Yaskawa INFORM job: 4043MM.JBI

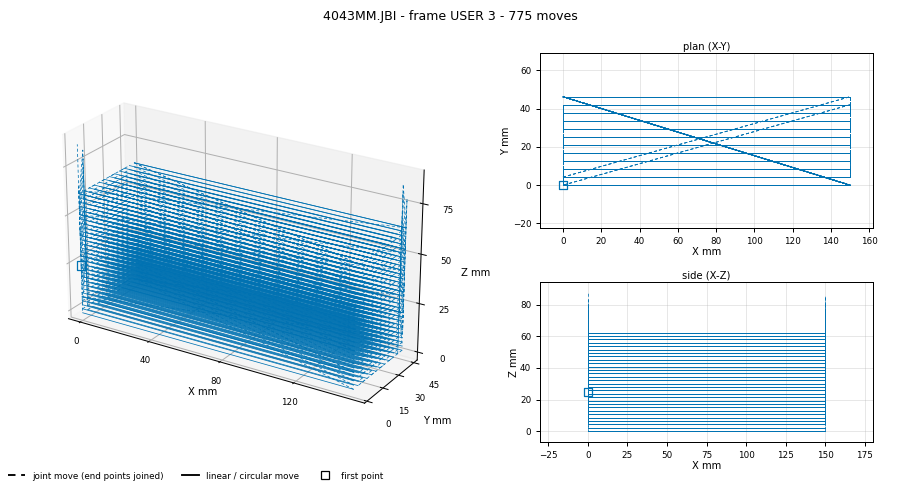
[picture p0: tool path of 4043MM.JBI in frame USER 3, 775 of 775 moves have a stored position in this frame; points joined in program order, loops and branches not executed]
/JOB
//NAME 4043MM
//POS
///NPOS 775,0,0,0,0,0
///USER 3
///TOOL 1
///POSTYPE USER
///RECTAN
///RCONF 1,0,0,0,0,0,0,0,0,0,0,0,0,0,0,0,0,0,0,0,0,0,0,0
C00000=0.000,0.000,25.000,0.0000,0.0000,-110.0000
C00001=0.000,0.000,0.000,0.0000,0.0000,-110.0000
C00002=150.000,0.000,0.000,0.0000,0.0000,-110.0000
C00003=0.000,46.200,0.000,0.0000,0.0000,-110.0000
C00004=150.000,46.200,0.000,0.0000,0.0000,-110.0000
C00005=150.000,4.200,0.000,0.0000,0.0000,-110.0000
C00006=0.000,4.200,0.000,0.0000,0.0000,-110.0000
C00007=0.000,8.400,0.000,0.0000,0.0000,-110.0000
C00008=150.000,8.400,0.000,0.0000,0.0000,-110.0000
C00009=150.000,12.600,0.000,0.0000,0.0000,-110.0000
C00010=0.000,12.600,0.000,0.0000,0.0000,-110.0000
C00011=0.000,16.800,0.000,0.0000,0.0000,-110.0000
C00012=150.000,16.800,0.000,0.0000,0.0000,-110.0000
C00013=150.000,21.000,0.000,0.0000,0.0000,-110.0000
C00014=0.000,21.000,0.000,0.0000,0.0000,-110.0000
C00015=0.000,25.200,0.000,0.0000,0.0000,-110.0000
C00016=150.000,25.200,0.000,0.0000,0.0000,-110.0000
C00017=150.000,29.400,0.000,0.0000,0.0000,-110.0000
C00018=0.000,29.400,0.000,0.0000,0.0000,-110.0000
C00019=0.000,33.600,0.000,0.0000,0.0000,-110.0000
C00020=150.000,33.600,0.000,0.0000,0.0000,-110.0000
C00021=150.000,37.800,0.000,0.0000,0.0000,-110.0000
C00022=0.000,37.800,0.000,0.0000,0.0000,-110.0000
C00023=0.000,42.000,0.000,0.0000,0.0000,-110.0000
C00024=150.000,42.000,0.000,0.0000,0.0000,-110.0000
C00025=150.000,42.000,25.000,0.0000,0.0000,-110.0000
C00026=150.000,46.200,2.150,0.0000,0.0000,-110.0000
C00027=0.000,46.200,2.150,0.0000,0.0000,-110.0000
C00028=150.000,0.000,2.150,0.0000,0.0000,-110.0000
C00029=0.000,0.000,2.150,0.0000,0.0000,-110.0000
C00030=0.000,42.000,2.150,0.0000,0.0000,-110.0000
C00031=150.000,42.000,2.150,0.0000,0.0000,-110.0000
C00032=150.000,37.800,2.150,0.0000,0.0000,-110.0000
C00033=0.000,37.800,2.150,0.0000,0.0000,-110.0000
C00034=0.000,33.600,2.150,0.0000,0.0000,-110.0000
C00035=150.000,33.600,2.150,0.0000,0.0000,-110.0000
C00036=150.000,29.400,2.150,0.0000,0.0000,-110.0000
C00037=0.000,29.400,2.150,0.0000,0.0000,-110.0000
C00038=0.000,25.200,2.150,0.0000,0.0000,-110.0000
C00039=150.000,25.200,2.150,0.0000,0.0000,-110.0000
C00040=150.000,21.000,2.150,0.0000,0.0000,-110.0000
C00041=0.000,21.000,2.150,0.0000,0.0000,-110.0000
C00042=0.000,16.800,2.150,0.0000,0.0000,-110.0000
C00043=150.000,16.800,2.150,0.0000,0.0000,-110.0000
C00044=150.000,12.600,2.150,0.0000,0.0000,-110.0000
C00045=0.000,12.600,2.150,0.0000,0.0000,-110.0000
C00046=0.000,8.400,2.150,0.0000,0.0000,-110.0000
C00047=150.000,8.400,2.150,0.0000,0.0000,-110.0000
C00048=150.000,4.200,2.150,0.0000,0.0000,-110.0000
C00049=0.000,4.200,2.150,0.0000,0.0000,-110.0000
C00050=0.000,4.200,27.150,0.0000,0.0000,-110.0000
C00051=0.000,0.000,4.300,0.0000,0.0000,-110.0000
C00052=150.000,0.000,4.300,0.0000,0.0000,-110.0000
C00053=0.000,46.200,4.300,0.0000,0.0000,-110.0000
C00054=150.000,46.200,4.300,0.0000,0.0000,-110.0000
C00055=150.000,4.200,4.300,0.0000,0.0000,-110.0000
C00056=0.000,4.200,4.300,0.0000,0.0000,-110.0000
C00057=0.000,8.400,4.300,0.0000,0.0000,-110.0000
C00058=150.000,8.400,4.300,0.0000,0.0000,-110.0000
C00059=150.000,12.600,4.300,0.0000,0.0000,-110.0000
C00060=0.000,12.600,4.300,0.0000,0.0000,-110.0000
C00061=0.000,16.800,4.300,0.0000,0.0000,-110.0000
C00062=150.000,16.800,4.300,0.0000,0.0000,-110.0000
C00063=150.000,21.000,4.300,0.0000,0.0000,-110.0000
C00064=0.000,21.000,4.300,0.0000,0.0000,-110.0000
C00065=0.000,25.200,4.300,0.0000,0.0000,-110.0000
C00066=150.000,25.200,4.300,0.0000,0.0000,-110.0000
C00067=150.000,29.400,4.300,0.0000,0.0000,-110.0000
C00068=0.000,29.400,4.300,0.0000,0.0000,-110.0000
C00069=0.000,33.600,4.300,0.0000,0.0000,-110.0000
C00070=150.000,33.600,4.300,0.0000,0.0000,-110.0000
C00071=150.000,37.800,4.300,0.0000,0.0000,-110.0000
C00072=0.000,37.800,4.300,0.0000,0.0000,-110.0000
C00073=0.000,42.000,4.300,0.0000,0.0000,-110.0000
C00074=150.000,42.000,4.300,0.0000,0.0000,-110.0000
C00075=150.000,42.000,29.300,0.0000,0.0000,-110.0000
C00076=150.000,46.200,6.450,0.0000,0.0000,-110.0000
C00077=0.000,46.200,6.450,0.0000,0.0000,-110.0000
C00078=150.000,0.000,6.450,0.0000,0.0000,-110.0000
C00079=0.000,0.000,6.450,0.0000,0.0000,-110.0000
C00080=0.000,42.000,6.450,0.0000,0.0000,-110.0000
C00081=150.000,42.000,6.450,0.0000,0.0000,-110.0000
C00082=150.000,37.800,6.450,0.0000,0.0000,-110.0000
C00083=0.000,37.800,6.450,0.0000,0.0000,-110.0000
C00084=0.000,33.600,6.450,0.0000,0.0000,-110.0000
C00085=150.000,33.600,6.450,0.0000,0.0000,-110.0000
C00086=150.000,29.400,6.450,0.0000,0.0000,-110.0000
C00087=0.000,29.400,6.450,0.0000,0.0000,-110.0000
C00088=0.000,25.200,6.450,0.0000,0.0000,-110.0000
C00089=150.000,25.200,6.450,0.0000,0.0000,-110.0000
C00090=150.000,21.000,6.450,0.0000,0.0000,-110.0000
C00091=0.000,21.000,6.450,0.0000,0.0000,-110.0000
C00092=0.000,16.800,6.450,0.0000,0.0000,-110.0000
C00093=150.000,16.800,6.450,0.0000,0.0000,-110.0000
C00094=150.000,12.600,6.450,0.0000,0.0000,-110.0000
C00095=0.000,12.600,6.450,0.0000,0.0000,-110.0000
C00096=0.000,8.400,6.450,0.0000,0.0000,-110.0000
C00097=150.000,8.400,6.450,0.0000,0.0000,-110.0000
C00098=150.000,4.200,6.450,0.0000,0.0000,-110.0000
C00099=0.000,4.200,6.450,0.0000,0.0000,-110.0000
C00100=0.000,4.200,31.450,0.0000,0.0000,-110.0000
C00101=0.000,0.000,8.600,0.0000,0.0000,-110.0000
C00102=150.000,0.000,8.600,0.0000,0.0000,-110.0000
C00103=0.000,46.200,8.600,0.0000,0.0000,-110.0000
C00104=150.000,46.200,8.600,0.0000,0.0000,-110.0000
C00105=150.000,4.200,8.600,0.0000,0.0000,-110.0000
C00106=0.000,4.200,8.600,0.0000,0.0000,-110.0000
C00107=0.000,8.400,8.600,0.0000,0.0000,-110.0000
C00108=150.000,8.400,8.600,0.0000,0.0000,-110.0000
C00109=150.000,12.600,8.600,0.0000,0.0000,-110.0000
C00110=0.000,12.600,8.600,0.0000,0.0000,-110.0000
C00111=0.000,16.800,8.600,0.0000,0.0000,-110.0000
C00112=150.000,16.800,8.600,0.0000,0.0000,-110.0000
C00113=150.000,21.000,8.600,0.0000,0.0000,-110.0000
C00114=0.000,21.000,8.600,0.0000,0.0000,-110.0000
C00115=0.000,25.200,8.600,0.0000,0.0000,-110.0000
C00116=150.000,25.200,8.600,0.0000,0.0000,-110.0000
C00117=150.000,29.400,8.600,0.0000,0.0000,-110.0000
C00118=0.000,29.400,8.600,0.0000,0.0000,-110.0000
C00119=0.000,33.600,8.600,0.0000,0.0000,-110.0000
C00120=150.000,33.600,8.600,0.0000,0.0000,-110.0000
C00121=150.000,37.800,8.600,0.0000,0.0000,-110.0000
C00122=0.000,37.800,8.600,0.0000,0.0000,-110.0000
C00123=0.000,42.000,8.600,0.0000,0.0000,-110.0000
C00124=150.000,42.000,8.600,0.0000,0.0000,-110.0000
C00125=0.000,0.000,8.600,0.0000,0.0000,-110.0000
C00126=150.000,0.000,8.600,0.0000,0.0000,-110.0000
C00127=0.000,46.200,8.600,0.0000,0.0000,-110.0000
C00128=150.000,46.200,8.600,0.0000,0.0000,-110.0000
C00129=150.000,46.200,33.600,0.0000,0.0000,-110.0000
C00130=150.000,46.200,10.750,0.0000,0.0000,-110.0000
C00131=0.000,46.200,10.750,0.0000,0.0000,-110.0000
C00132=150.000,0.000,10.750,0.0000,0.0000,-110.0000
C00133=0.000,0.000,10.750,0.0000,0.0000,-110.0000
C00134=0.000,42.000,10.750,0.0000,0.0000,-110.0000
C00135=150.000,42.000,10.750,0.0000,0.0000,-110.0000
C00136=150.000,37.800,10.750,0.0000,0.0000,-110.0000
C00137=0.000,37.800,10.750,0.0000,0.0000,-110.0000
C00138=0.000,33.600,10.750,0.0000,0.0000,-110.0000
C00139=150.000,33.600,10.750,0.0000,0.0000,-110.0000
C00140=150.000,29.400,10.750,0.0000,0.0000,-110.0000
C00141=0.000,29.400,10.750,0.0000,0.0000,-110.0000
C00142=0.000,25.200,10.750,0.0000,0.0000,-110.0000
C00143=150.000,25.200,10.750,0.0000,0.0000,-110.0000
C00144=150.000,21.000,10.750,0.0000,0.0000,-110.0000
C00145=0.000,21.000,10.750,0.0000,0.0000,-110.0000
C00146=0.000,16.800,10.750,0.0000,0.0000,-110.0000
C00147=150.000,16.800,10.750,0.0000,0.0000,-110.0000
C00148=150.000,12.600,10.750,0.0000,0.0000,-110.0000
C00149=0.000,12.600,10.750,0.0000,0.0000,-110.0000
C00150=0.000,8.400,10.750,0.0000,0.0000,-110.0000
C00151=150.000,8.400,10.750,0.0000,0.0000,-110.0000
C00152=150.000,4.200,10.750,0.0000,0.0000,-110.0000
C00153=0.000,4.200,10.750,0.0000,0.0000,-110.0000
C00154=0.000,4.200,35.750,0.0000,0.0000,-110.0000
C00155=0.000,0.000,12.900,0.0000,0.0000,-110.0000
C00156=150.000,0.000,12.900,0.0000,0.0000,-110.0000
C00157=0.000,46.200,12.900,0.0000,0.0000,-110.0000
C00158=150.000,46.200,12.900,0.0000,0.0000,-110.0000
C00159=150.000,4.200,12.900,0.0000,0.0000,-110.0000
C00160=0.000,4.200,12.900,0.0000,0.0000,-110.0000
C00161=0.000,8.400,12.900,0.0000,0.0000,-110.0000
C00162=150.000,8.400,12.900,0.0000,0.0000,-110.0000
C00163=150.000,12.600,12.900,0.0000,0.0000,-110.0000
C00164=0.000,12.600,12.900,0.0000,0.0000,-110.0000
C00165=0.000,16.800,12.900,0.0000,0.0000,-110.0000
C00166=150.000,16.800,12.900,0.0000,0.0000,-110.0000
C00167=150.000,21.000,12.900,0.0000,0.0000,-110.0000
C00168=0.000,21.000,12.900,0.0000,0.0000,-110.0000
C00169=0.000,25.200,12.900,0.0000,0.0000,-110.0000
C00170=150.000,25.200,12.900,0.0000,0.0000,-110.0000
C00171=150.000,29.400,12.900,0.0000,0.0000,-110.0000
C00172=0.000,29.400,12.900,0.0000,0.0000,-110.0000
C00173=0.000,33.600,12.900,0.0000,0.0000,-110.0000
C00174=150.000,33.600,12.900,0.0000,0.0000,-110.0000
C00175=150.000,37.800,12.900,0.0000,0.0000,-110.0000
C00176=0.000,37.800,12.900,0.0000,0.0000,-110.0000
C00177=0.000,42.000,12.900,0.0000,0.0000,-110.0000
C00178=150.000,42.000,12.900,0.0000,0.0000,-110.0000
C00179=150.000,42.000,37.900,0.0000,0.0000,-110.0000
C00180=150.000,46.200,15.050,0.0000,0.0000,-110.0000
C00181=0.000,46.200,15.050,0.0000,0.0000,-110.0000
C00182=150.000,0.000,15.050,0.0000,0.0000,-110.0000
C00183=0.000,0.000,15.050,0.0000,0.0000,-110.0000
C00184=0.000,42.000,15.050,0.0000,0.0000,-110.0000
C00185=150.000,42.000,15.050,0.0000,0.0000,-110.0000
C00186=150.000,37.800,15.050,0.0000,0.0000,-110.0000
C00187=0.000,37.800,15.050,0.0000,0.0000,-110.0000
C00188=0.000,33.600,15.050,0.0000,0.0000,-110.0000
C00189=150.000,33.600,15.050,0.0000,0.0000,-110.0000
C00190=150.000,29.400,15.050,0.0000,0.0000,-110.0000
C00191=0.000,29.400,15.050,0.0000,0.0000,-110.0000
C00192=0.000,25.200,15.050,0.0000,0.0000,-110.0000
C00193=150.000,25.200,15.050,0.0000,0.0000,-110.0000
C00194=150.000,21.000,15.050,0.0000,0.0000,-110.0000
C00195=0.000,21.000,15.050,0.0000,0.0000,-110.0000
C00196=0.000,16.800,15.050,0.0000,0.0000,-110.0000
C00197=150.000,16.800,15.050,0.0000,0.0000,-110.0000
C00198=150.000,12.600,15.050,0.0000,0.0000,-110.0000
C00199=0.000,12.600,15.050,0.0000,0.0000,-110.0000
C00200=0.000,8.400,15.050,0.0000,0.0000,-110.0000
C00201=150.000,8.400,15.050,0.0000,0.0000,-110.0000
C00202=150.000,4.200,15.050,0.0000,0.0000,-110.0000
C00203=0.000,4.200,15.050,0.0000,0.0000,-110.0000
C00204=0.000,4.200,40.050,0.0000,0.0000,-110.0000
C00205=0.000,0.000,17.200,0.0000,0.0000,-110.0000
C00206=150.000,0.000,17.200,0.0000,0.0000,-110.0000
C00207=0.000,46.200,17.200,0.0000,0.0000,-110.0000
C00208=150.000,46.200,17.200,0.0000,0.0000,-110.0000
C00209=150.000,4.200,17.200,0.0000,0.0000,-110.0000
C00210=0.000,4.200,17.200,0.0000,0.0000,-110.0000
C00211=0.000,8.400,17.200,0.0000,0.0000,-110.0000
C00212=150.000,8.400,17.200,0.0000,0.0000,-110.0000
C00213=150.000,12.600,17.200,0.0000,0.0000,-110.0000
C00214=0.000,12.600,17.200,0.0000,0.0000,-110.0000
C00215=0.000,16.800,17.200,0.0000,0.0000,-110.0000
C00216=150.000,16.800,17.200,0.0000,0.0000,-110.0000
C00217=150.000,21.000,17.200,0.0000,0.0000,-110.0000
C00218=0.000,21.000,17.200,0.0000,0.0000,-110.0000
C00219=0.000,25.200,17.200,0.0000,0.0000,-110.0000
C00220=150.000,25.200,17.200,0.0000,0.0000,-110.0000
C00221=150.000,29.400,17.200,0.0000,0.0000,-110.0000
C00222=0.000,29.400,17.200,0.0000,0.0000,-110.0000
C00223=0.000,33.600,17.200,0.0000,0.0000,-110.0000
C00224=150.000,33.600,17.200,0.0000,0.0000,-110.0000
C00225=150.000,37.800,17.200,0.0000,0.0000,-110.0000
C00226=0.000,37.800,17.200,0.0000,0.0000,-110.0000
C00227=0.000,42.000,17.200,0.0000,0.0000,-110.0000
C00228=150.000,42.000,17.200,0.0000,0.0000,-110.0000
C00229=150.000,42.000,42.200,0.0000,0.0000,-110.0000
C00230=150.000,46.200,19.350,0.0000,0.0000,-110.0000
C00231=0.000,46.200,19.350,0.0000,0.0000,-110.0000
C00232=150.000,0.000,19.350,0.0000,0.0000,-110.0000
C00233=0.000,0.000,19.350,0.0000,0.0000,-110.0000
C00234=0.000,42.000,19.350,0.0000,0.0000,-110.0000
C00235=150.000,42.000,19.350,0.0000,0.0000,-110.0000
C00236=150.000,37.800,19.350,0.0000,0.0000,-110.0000
C00237=0.000,37.800,19.350,0.0000,0.0000,-110.0000
C00238=0.000,33.600,19.350,0.0000,0.0000,-110.0000
C00239=150.000,33.600,19.350,0.0000,0.0000,-110.0000
C00240=150.000,29.400,19.350,0.0000,0.0000,-110.0000
C00241=0.000,29.400,19.350,0.0000,0.0000,-110.0000
C00242=0.000,25.200,19.350,0.0000,0.0000,-110.0000
C00243=150.000,25.200,19.350,0.0000,0.0000,-110.0000
C00244=150.000,21.000,19.350,0.0000,0.0000,-110.0000
C00245=0.000,21.000,19.350,0.0000,0.0000,-110.0000
C00246=0.000,16.800,19.350,0.0000,0.0000,-110.0000
C00247=150.000,16.800,19.350,0.0000,0.0000,-110.0000
C00248=150.000,12.600,19.350,0.0000,0.0000,-110.0000
C00249=0.000,12.600,19.350,0.0000,0.0000,-110.0000
C00250=0.000,8.400,19.350,0.0000,0.0000,-110.0000
C00251=150.000,8.400,19.350,0.0000,0.0000,-110.0000
C00252=150.000,4.200,19.350,0.0000,0.0000,-110.0000
C00253=0.000,4.200,19.350,0.0000,0.0000,-110.0000
C00254=150.000,46.200,19.350,0.0000,0.0000,-110.0000
C00255=0.000,46.200,19.350,0.0000,0.0000,-110.0000
C00256=150.000,0.000,19.350,0.0000,0.0000,-110.0000
C00257=0.000,0.000,19.350,0.0000,0.0000,-110.0000
C00258=0.000,0.000,44.350,0.0000,0.0000,-110.0000
C00259=0.000,0.000,21.500,0.0000,0.0000,-110.0000
C00260=150.000,0.000,21.500,0.0000,0.0000,-110.0000
C00261=0.000,46.200,21.500,0.0000,0.0000,-110.0000
C00262=150.000,46.200,21.500,0.0000,0.0000,-110.0000
C00263=150.000,4.200,21.500,0.0000,0.0000,-110.0000
C00264=0.000,4.200,21.500,0.0000,0.0000,-110.0000
C00265=0.000,8.400,21.500,0.0000,0.0000,-110.0000
C00266=150.000,8.400,21.500,0.0000,0.0000,-110.0000
C00267=150.000,12.600,21.500,0.0000,0.0000,-110.0000
C00268=0.000,12.600,21.500,0.0000,0.0000,-110.0000
C00269=0.000,16.800,21.500,0.0000,0.0000,-110.0000
C00270=150.000,16.800,21.500,0.0000,0.0000,-110.0000
C00271=150.000,21.000,21.500,0.0000,0.0000,-110.0000
C00272=0.000,21.000,21.500,0.0000,0.0000,-110.0000
C00273=0.000,25.200,21.500,0.0000,0.0000,-110.0000
C00274=150.000,25.200,21.500,0.0000,0.0000,-110.0000
C00275=150.000,29.400,21.500,0.0000,0.0000,-110.0000
C00276=0.000,29.400,21.500,0.0000,0.0000,-110.0000
C00277=0.000,33.600,21.500,0.0000,0.0000,-110.0000
C00278=150.000,33.600,21.500,0.0000,0.0000,-110.0000
C00279=150.000,37.800,21.500,0.0000,0.0000,-110.0000
C00280=0.000,37.800,21.500,0.0000,0.0000,-110.0000
C00281=0.000,42.000,21.500,0.0000,0.0000,-110.0000
C00282=150.000,42.000,21.500,0.0000,0.0000,-110.0000
C00283=150.000,42.000,46.500,0.0000,0.0000,-110.0000
C00284=150.000,46.200,23.650,0.0000,0.0000,-110.0000
C00285=0.000,46.200,23.650,0.0000,0.0000,-110.0000
C00286=150.000,0.000,23.650,0.0000,0.0000,-110.0000
C00287=0.000,0.000,23.650,0.0000,0.0000,-110.0000
C00288=0.000,42.000,23.650,0.0000,0.0000,-110.0000
C00289=150.000,42.000,23.650,0.0000,0.0000,-110.0000
C00290=150.000,37.800,23.650,0.0000,0.0000,-110.0000
C00291=0.000,37.800,23.650,0.0000,0.0000,-110.0000
C00292=0.000,33.600,23.650,0.0000,0.0000,-110.0000
C00293=150.000,33.600,23.650,0.0000,0.0000,-110.0000
C00294=150.000,29.400,23.650,0.0000,0.0000,-110.0000
C00295=0.000,29.400,23.650,0.0000,0.0000,-110.0000
C00296=0.000,25.200,23.650,0.0000,0.0000,-110.0000
C00297=150.000,25.200,23.650,0.0000,0.0000,-110.0000
C00298=150.000,21.000,23.650,0.0000,0.0000,-110.0000
C00299=0.000,21.000,23.650,0.0000,0.0000,-110.0000
C00300=0.000,16.800,23.650,0.0000,0.0000,-110.0000
C00301=150.000,16.800,23.650,0.0000,0.0000,-110.0000
C00302=150.000,12.600,23.650,0.0000,0.0000,-110.0000
C00303=0.000,12.600,23.650,0.0000,0.0000,-110.0000
C00304=0.000,8.400,23.650,0.0000,0.0000,-110.0000
C00305=150.000,8.400,23.650,0.0000,0.0000,-110.0000
C00306=150.000,4.200,23.650,0.0000,0.0000,-110.0000
C00307=0.000,4.200,23.650,0.0000,0.0000,-110.0000
C00308=0.000,4.200,48.650,0.0000,0.0000,-110.0000
C00309=0.000,0.000,25.800,0.0000,0.0000,-110.0000
C00310=150.000,0.000,25.800,0.0000,0.0000,-110.0000
C00311=0.000,46.200,25.800,0.0000,0.0000,-110.0000
C00312=150.000,46.200,25.800,0.0000,0.0000,-110.0000
C00313=150.000,4.200,25.800,0.0000,0.0000,-110.0000
C00314=0.000,4.200,25.800,0.0000,0.0000,-110.0000
C00315=0.000,8.400,25.800,0.0000,0.0000,-110.0000
C00316=150.000,8.400,25.800,0.0000,0.0000,-110.0000
C00317=150.000,12.600,25.800,0.0000,0.0000,-110.0000
C00318=0.000,12.600,25.800,0.0000,0.0000,-110.0000
C00319=0.000,16.800,25.800,0.0000,0.0000,-110.0000
C00320=150.000,16.800,25.800,0.0000,0.0000,-110.0000
C00321=150.000,21.000,25.800,0.0000,0.0000,-110.0000
C00322=0.000,21.000,25.800,0.0000,0.0000,-110.0000
C00323=0.000,25.200,25.800,0.0000,0.0000,-110.0000
C00324=150.000,25.200,25.800,0.0000,0.0000,-110.0000
C00325=150.000,29.400,25.800,0.0000,0.0000,-110.0000
C00326=0.000,29.400,25.800,0.0000,0.0000,-110.0000
C00327=0.000,33.600,25.800,0.0000,0.0000,-110.0000
C00328=150.000,33.600,25.800,0.0000,0.0000,-110.0000
C00329=150.000,37.800,25.800,0.0000,0.0000,-110.0000
C00330=0.000,37.800,25.800,0.0000,0.0000,-110.0000
C00331=0.000,42.000,25.800,0.0000,0.0000,-110.0000
C00332=150.000,42.000,25.800,0.0000,0.0000,-110.0000
C00333=150.000,42.000,50.800,0.0000,0.0000,-110.0000
C00334=150.000,46.200,27.950,0.0000,0.0000,-110.0000
C00335=0.000,46.200,27.950,0.0000,0.0000,-110.0000
C00336=150.000,0.000,27.950,0.0000,0.0000,-110.0000
C00337=0.000,0.000,27.950,0.0000,0.0000,-110.0000
C00338=0.000,42.000,27.950,0.0000,0.0000,-110.0000
C00339=150.000,42.000,27.950,0.0000,0.0000,-110.0000
C00340=150.000,37.800,27.950,0.0000,0.0000,-110.0000
C00341=0.000,37.800,27.950,0.0000,0.0000,-110.0000
C00342=0.000,33.600,27.950,0.0000,0.0000,-110.0000
C00343=150.000,33.600,27.950,0.0000,0.0000,-110.0000
C00344=150.000,29.400,27.950,0.0000,0.0000,-110.0000
C00345=0.000,29.400,27.950,0.0000,0.0000,-110.0000
C00346=0.000,25.200,27.950,0.0000,0.0000,-110.0000
C00347=150.000,25.200,27.950,0.0000,0.0000,-110.0000
C00348=150.000,21.000,27.950,0.0000,0.0000,-110.0000
C00349=0.000,21.000,27.950,0.0000,0.0000,-110.0000
C00350=0.000,16.800,27.950,0.0000,0.0000,-110.0000
C00351=150.000,16.800,27.950,0.0000,0.0000,-110.0000
C00352=150.000,12.600,27.950,0.0000,0.0000,-110.0000
C00353=0.000,12.600,27.950,0.0000,0.0000,-110.0000
C00354=0.000,8.400,27.950,0.0000,0.0000,-110.0000
C00355=150.000,8.400,27.950,0.0000,0.0000,-110.0000
C00356=150.000,4.200,27.950,0.0000,0.0000,-110.0000
C00357=0.000,4.200,27.950,0.0000,0.0000,-110.0000
C00358=0.000,4.200,52.950,0.0000,0.0000,-110.0000
C00359=0.000,0.000,30.100,0.0000,0.0000,-110.0000
C00360=150.000,0.000,30.100,0.0000,0.0000,-110.0000
C00361=0.000,46.200,30.100,0.0000,0.0000,-110.0000
C00362=150.000,46.200,30.100,0.0000,0.0000,-110.0000
C00363=150.000,4.200,30.100,0.0000,0.0000,-110.0000
C00364=0.000,4.200,30.100,0.0000,0.0000,-110.0000
C00365=0.000,8.400,30.100,0.0000,0.0000,-110.0000
C00366=150.000,8.400,30.100,0.0000,0.0000,-110.0000
C00367=150.000,12.600,30.100,0.0000,0.0000,-110.0000
C00368=0.000,12.600,30.100,0.0000,0.0000,-110.0000
C00369=0.000,16.800,30.100,0.0000,0.0000,-110.0000
C00370=150.000,16.800,30.100,0.0000,0.0000,-110.0000
C00371=150.000,21.000,30.100,0.0000,0.0000,-110.0000
C00372=0.000,21.000,30.100,0.0000,0.0000,-110.0000
C00373=0.000,25.200,30.100,0.0000,0.0000,-110.0000
C00374=150.000,25.200,30.100,0.0000,0.0000,-110.0000
C00375=150.000,29.400,30.100,0.0000,0.0000,-110.0000
C00376=0.000,29.400,30.100,0.0000,0.0000,-110.0000
C00377=0.000,33.600,30.100,0.0000,0.0000,-110.0000
C00378=150.000,33.600,30.100,0.0000,0.0000,-110.0000
C00379=150.000,37.800,30.100,0.0000,0.0000,-110.0000
C00380=0.000,37.800,30.100,0.0000,0.0000,-110.0000
C00381=0.000,42.000,30.100,0.0000,0.0000,-110.0000
C00382=150.000,42.000,30.100,0.0000,0.0000,-110.0000
C00383=0.000,0.000,30.100,0.0000,0.0000,-110.0000
C00384=150.000,0.000,30.100,0.0000,0.0000,-110.0000
C00385=0.000,46.200,30.100,0.0000,0.0000,-110.0000
C00386=150.000,46.200,30.100,0.0000,0.0000,-110.0000
C00387=150.000,46.200,55.100,0.0000,0.0000,-110.0000
C00388=150.000,46.200,32.250,0.0000,0.0000,-110.0000
C00389=0.000,46.200,32.250,0.0000,0.0000,-110.0000
C00390=150.000,0.000,32.250,0.0000,0.0000,-110.0000
C00391=0.000,0.000,32.250,0.0000,0.0000,-110.0000
C00392=0.000,42.000,32.250,0.0000,0.0000,-110.0000
C00393=150.000,42.000,32.250,0.0000,0.0000,-110.0000
C00394=150.000,37.800,32.250,0.0000,0.0000,-110.0000
C00395=0.000,37.800,32.250,0.0000,0.0000,-110.0000
C00396=0.000,33.600,32.250,0.0000,0.0000,-110.0000
C00397=150.000,33.600,32.250,0.0000,0.0000,-110.0000
C00398=150.000,29.400,32.250,0.0000,0.0000,-110.0000
C00399=0.000,29.400,32.250,0.0000,0.0000,-110.0000
C00400=0.000,25.200,32.250,0.0000,0.0000,-110.0000
C00401=150.000,25.200,32.250,0.0000,0.0000,-110.0000
C00402=150.000,21.000,32.250,0.0000,0.0000,-110.0000
C00403=0.000,21.000,32.250,0.0000,0.0000,-110.0000
C00404=0.000,16.800,32.250,0.0000,0.0000,-110.0000
C00405=150.000,16.800,32.250,0.0000,0.0000,-110.0000
C00406=150.000,12.600,32.250,0.0000,0.0000,-110.0000
C00407=0.000,12.600,32.250,0.0000,0.0000,-110.0000
C00408=0.000,8.400,32.250,0.0000,0.0000,-110.0000
C00409=150.000,8.400,32.250,0.0000,0.0000,-110.0000
C00410=150.000,4.200,32.250,0.0000,0.0000,-110.0000
C00411=0.000,4.200,32.250,0.0000,0.0000,-110.0000
C00412=0.000,4.200,57.250,0.0000,0.0000,-110.0000
C00413=0.000,0.000,34.400,0.0000,0.0000,-110.0000
C00414=150.000,0.000,34.400,0.0000,0.0000,-110.0000
C00415=0.000,46.200,34.400,0.0000,0.0000,-110.0000
C00416=150.000,46.200,34.400,0.0000,0.0000,-110.0000
C00417=150.000,4.200,34.400,0.0000,0.0000,-110.0000
C00418=0.000,4.200,34.400,0.0000,0.0000,-110.0000
C00419=0.000,8.400,34.400,0.0000,0.0000,-110.0000
C00420=150.000,8.400,34.400,0.0000,0.0000,-110.0000
C00421=150.000,12.600,34.400,0.0000,0.0000,-110.0000
C00422=0.000,12.600,34.400,0.0000,0.0000,-110.0000
C00423=0.000,16.800,34.400,0.0000,0.0000,-110.0000
C00424=150.000,16.800,34.400,0.0000,0.0000,-110.0000
C00425=150.000,21.000,34.400,0.0000,0.0000,-110.0000
C00426=0.000,21.000,34.400,0.0000,0.0000,-110.0000
C00427=0.000,25.200,34.400,0.0000,0.0000,-110.0000
C00428=150.000,25.200,34.400,0.0000,0.0000,-110.0000
C00429=150.000,29.400,34.400,0.0000,0.0000,-110.0000
C00430=0.000,29.400,34.400,0.0000,0.0000,-110.0000
C00431=0.000,33.600,34.400,0.0000,0.0000,-110.0000
C00432=150.000,33.600,34.400,0.0000,0.0000,-110.0000
C00433=150.000,37.800,34.400,0.0000,0.0000,-110.0000
C00434=0.000,37.800,34.400,0.0000,0.0000,-110.0000
C00435=0.000,42.000,34.400,0.0000,0.0000,-110.0000
C00436=150.000,42.000,34.400,0.0000,0.0000,-110.0000
C00437=150.000,42.000,59.400,0.0000,0.0000,-110.0000
C00438=150.000,46.200,36.550,0.0000,0.0000,-110.0000
C00439=0.000,46.200,36.550,0.0000,0.0000,-110.0000
C00440=150.000,0.000,36.550,0.0000,0.0000,-110.0000
C00441=0.000,0.000,36.550,0.0000,0.0000,-110.0000
C00442=0.000,42.000,36.550,0.0000,0.0000,-110.0000
C00443=150.000,42.000,36.550,0.0000,0.0000,-110.0000
C00444=150.000,37.800,36.550,0.0000,0.0000,-110.0000
C00445=0.000,37.800,36.550,0.0000,0.0000,-110.0000
C00446=0.000,33.600,36.550,0.0000,0.0000,-110.0000
C00447=150.000,33.600,36.550,0.0000,0.0000,-110.0000
C00448=150.000,29.400,36.550,0.0000,0.0000,-110.0000
C00449=0.000,29.400,36.550,0.0000,0.0000,-110.0000
C00450=0.000,25.200,36.550,0.0000,0.0000,-110.0000
C00451=150.000,25.200,36.550,0.0000,0.0000,-110.0000
C00452=150.000,21.000,36.550,0.0000,0.0000,-110.0000
C00453=0.000,21.000,36.550,0.0000,0.0000,-110.0000
C00454=0.000,16.800,36.550,0.0000,0.0000,-110.0000
C00455=150.000,16.800,36.550,0.0000,0.0000,-110.0000
C00456=150.000,12.600,36.550,0.0000,0.0000,-110.0000
C00457=0.000,12.600,36.550,0.0000,0.0000,-110.0000
C00458=0.000,8.400,36.550,0.0000,0.0000,-110.0000
C00459=150.000,8.400,36.550,0.0000,0.0000,-110.0000
C00460=150.000,4.200,36.550,0.0000,0.0000,-110.0000
C00461=0.000,4.200,36.550,0.0000,0.0000,-110.0000
C00462=0.000,4.200,61.550,0.0000,0.0000,-110.0000
C00463=0.000,0.000,38.700,0.0000,0.0000,-110.0000
C00464=150.000,0.000,38.700,0.0000,0.0000,-110.0000
C00465=0.000,46.200,38.700,0.0000,0.0000,-110.0000
C00466=150.000,46.200,38.700,0.0000,0.0000,-110.0000
C00467=150.000,4.200,38.700,0.0000,0.0000,-110.0000
C00468=0.000,4.200,38.700,0.0000,0.0000,-110.0000
C00469=0.000,8.400,38.700,0.0000,0.0000,-110.0000
C00470=150.000,8.400,38.700,0.0000,0.0000,-110.0000
C00471=150.000,12.600,38.700,0.0000,0.0000,-110.0000
C00472=0.000,12.600,38.700,0.0000,0.0000,-110.0000
C00473=0.000,16.800,38.700,0.0000,0.0000,-110.0000
C00474=150.000,16.800,38.700,0.0000,0.0000,-110.0000
C00475=150.000,21.000,38.700,0.0000,0.0000,-110.0000
C00476=0.000,21.000,38.700,0.0000,0.0000,-110.0000
C00477=0.000,25.200,38.700,0.0000,0.0000,-110.0000
C00478=150.000,25.200,38.700,0.0000,0.0000,-110.0000
C00479=150.000,29.400,38.700,0.0000,0.0000,-110.0000
C00480=0.000,29.400,38.700,0.0000,0.0000,-110.0000
C00481=0.000,33.600,38.700,0.0000,0.0000,-110.0000
C00482=150.000,33.600,38.700,0.0000,0.0000,-110.0000
C00483=150.000,37.800,38.700,0.0000,0.0000,-110.0000
C00484=0.000,37.800,38.700,0.0000,0.0000,-110.0000
C00485=0.000,42.000,38.700,0.0000,0.0000,-110.0000
C00486=150.000,42.000,38.700,0.0000,0.0000,-110.0000
C00487=150.000,42.000,63.700,0.0000,0.0000,-110.0000
C00488=150.000,46.200,40.850,0.0000,0.0000,-110.0000
C00489=0.000,46.200,40.850,0.0000,0.0000,-110.0000
C00490=150.000,0.000,40.850,0.0000,0.0000,-110.0000
C00491=0.000,0.000,40.850,0.0000,0.0000,-110.0000
C00492=0.000,42.000,40.850,0.0000,0.0000,-110.0000
C00493=150.000,42.000,40.850,0.0000,0.0000,-110.0000
C00494=150.000,37.800,40.850,0.0000,0.0000,-110.0000
C00495=0.000,37.800,40.850,0.0000,0.0000,-110.0000
C00496=0.000,33.600,40.850,0.0000,0.0000,-110.0000
C00497=150.000,33.600,40.850,0.0000,0.0000,-110.0000
C00498=150.000,29.400,40.850,0.0000,0.0000,-110.0000
C00499=0.000,29.400,40.850,0.0000,0.0000,-110.0000
C00500=0.000,25.200,40.850,0.0000,0.0000,-110.0000
C00501=150.000,25.200,40.850,0.0000,0.0000,-110.0000
C00502=150.000,21.000,40.850,0.0000,0.0000,-110.0000
C00503=0.000,21.000,40.850,0.0000,0.0000,-110.0000
C00504=0.000,16.800,40.850,0.0000,0.0000,-110.0000
C00505=150.000,16.800,40.850,0.0000,0.0000,-110.0000
C00506=150.000,12.600,40.850,0.0000,0.0000,-110.0000
C00507=0.000,12.600,40.850,0.0000,0.0000,-110.0000
C00508=0.000,8.400,40.850,0.0000,0.0000,-110.0000
C00509=150.000,8.400,40.850,0.0000,0.0000,-110.0000
C00510=150.000,4.200,40.850,0.0000,0.0000,-110.0000
C00511=0.000,4.200,40.850,0.0000,0.0000,-110.0000
C00512=150.000,46.200,40.850,0.0000,0.0000,-110.0000
C00513=0.000,46.200,40.850,0.0000,0.0000,-110.0000
C00514=150.000,0.000,40.850,0.0000,0.0000,-110.0000
C00515=0.000,0.000,40.850,0.0000,0.0000,-110.0000
C00516=0.000,0.000,65.850,0.0000,0.0000,-110.0000
C00517=0.000,0.000,43.000,0.0000,0.0000,-110.0000
C00518=150.000,0.000,43.000,0.0000,0.0000,-110.0000
C00519=0.000,46.200,43.000,0.0000,0.0000,-110.0000
C00520=150.000,46.200,43.000,0.0000,0.0000,-110.0000
C00521=150.000,4.200,43.000,0.0000,0.0000,-110.0000
C00522=0.000,4.200,43.000,0.0000,0.0000,-110.0000
C00523=0.000,8.400,43.000,0.0000,0.0000,-110.0000
C00524=150.000,8.400,43.000,0.0000,0.0000,-110.0000
C00525=150.000,12.600,43.000,0.0000,0.0000,-110.0000
C00526=0.000,12.600,43.000,0.0000,0.0000,-110.0000
C00527=0.000,16.800,43.000,0.0000,0.0000,-110.0000
C00528=150.000,16.800,43.000,0.0000,0.0000,-110.0000
C00529=150.000,21.000,43.000,0.0000,0.0000,-110.0000
C00530=0.000,21.000,43.000,0.0000,0.0000,-110.0000
C00531=0.000,25.200,43.000,0.0000,0.0000,-110.0000
C00532=150.000,25.200,43.000,0.0000,0.0000,-110.0000
C00533=150.000,29.400,43.000,0.0000,0.0000,-110.0000
C00534=0.000,29.400,43.000,0.0000,0.0000,-110.0000
C00535=0.000,33.600,43.000,0.0000,0.0000,-110.0000
C00536=150.000,33.600,43.000,0.0000,0.0000,-110.0000
C00537=150.000,37.800,43.000,0.0000,0.0000,-110.0000
C00538=0.000,37.800,43.000,0.0000,0.0000,-110.0000
C00539=0.000,42.000,43.000,0.0000,0.0000,-110.0000
C00540=150.000,42.000,43.000,0.0000,0.0000,-110.0000
C00541=150.000,42.000,68.000,0.0000,0.0000,-110.0000
C00542=150.000,46.200,45.150,0.0000,0.0000,-110.0000
C00543=0.000,46.200,45.150,0.0000,0.0000,-110.0000
C00544=150.000,0.000,45.150,0.0000,0.0000,-110.0000
C00545=0.000,0.000,45.150,0.0000,0.0000,-110.0000
C00546=0.000,42.000,45.150,0.0000,0.0000,-110.0000
C00547=150.000,42.000,45.150,0.0000,0.0000,-110.0000
C00548=150.000,37.800,45.150,0.0000,0.0000,-110.0000
C00549=0.000,37.800,45.150,0.0000,0.0000,-110.0000
C00550=0.000,33.600,45.150,0.0000,0.0000,-110.0000
C00551=150.000,33.600,45.150,0.0000,0.0000,-110.0000
C00552=150.000,29.400,45.150,0.0000,0.0000,-110.0000
C00553=0.000,29.400,45.150,0.0000,0.0000,-110.0000
C00554=0.000,25.200,45.150,0.0000,0.0000,-110.0000
C00555=150.000,25.200,45.150,0.0000,0.0000,-110.0000
C00556=150.000,21.000,45.150,0.0000,0.0000,-110.0000
C00557=0.000,21.000,45.150,0.0000,0.0000,-110.0000
C00558=0.000,16.800,45.150,0.0000,0.0000,-110.0000
C00559=150.000,16.800,45.150,0.0000,0.0000,-110.0000
C00560=150.000,12.600,45.150,0.0000,0.0000,-110.0000
C00561=0.000,12.600,45.150,0.0000,0.0000,-110.0000
C00562=0.000,8.400,45.150,0.0000,0.0000,-110.0000
C00563=150.000,8.400,45.150,0.0000,0.0000,-110.0000
C00564=150.000,4.200,45.150,0.0000,0.0000,-110.0000
C00565=0.000,4.200,45.150,0.0000,0.0000,-110.0000
C00566=0.000,4.200,70.150,0.0000,0.0000,-110.0000
C00567=0.000,0.000,47.300,0.0000,0.0000,-110.0000
C00568=150.000,0.000,47.300,0.0000,0.0000,-110.0000
C00569=0.000,46.200,47.300,0.0000,0.0000,-110.0000
C00570=150.000,46.200,47.300,0.0000,0.0000,-110.0000
C00571=150.000,4.200,47.300,0.0000,0.0000,-110.0000
C00572=0.000,4.200,47.300,0.0000,0.0000,-110.0000
C00573=0.000,8.400,47.300,0.0000,0.0000,-110.0000
C00574=150.000,8.400,47.300,0.0000,0.0000,-110.0000
C00575=150.000,12.600,47.300,0.0000,0.0000,-110.0000
C00576=0.000,12.600,47.300,0.0000,0.0000,-110.0000
C00577=0.000,16.800,47.300,0.0000,0.0000,-110.0000
C00578=150.000,16.800,47.300,0.0000,0.0000,-110.0000
C00579=150.000,21.000,47.300,0.0000,0.0000,-110.0000
C00580=0.000,21.000,47.300,0.0000,0.0000,-110.0000
C00581=0.000,25.200,47.300,0.0000,0.0000,-110.0000
C00582=150.000,25.200,47.300,0.0000,0.0000,-110.0000
C00583=150.000,29.400,47.300,0.0000,0.0000,-110.0000
C00584=0.000,29.400,47.300,0.0000,0.0000,-110.0000
C00585=0.000,33.600,47.300,0.0000,0.0000,-110.0000
C00586=150.000,33.600,47.300,0.0000,0.0000,-110.0000
C00587=150.000,37.800,47.300,0.0000,0.0000,-110.0000
C00588=0.000,37.800,47.300,0.0000,0.0000,-110.0000
C00589=0.000,42.000,47.300,0.0000,0.0000,-110.0000
C00590=150.000,42.000,47.300,0.0000,0.0000,-110.0000
C00591=150.000,42.000,72.300,0.0000,0.0000,-110.0000
C00592=150.000,46.200,49.450,0.0000,0.0000,-110.0000
C00593=0.000,46.200,49.450,0.0000,0.0000,-110.0000
C00594=150.000,0.000,49.450,0.0000,0.0000,-110.0000
C00595=0.000,0.000,49.450,0.0000,0.0000,-110.0000
C00596=0.000,42.000,49.450,0.0000,0.0000,-110.0000
C00597=150.000,42.000,49.450,0.0000,0.0000,-110.0000
C00598=150.000,37.800,49.450,0.0000,0.0000,-110.0000
C00599=0.000,37.800,49.450,0.0000,0.0000,-110.0000
C00600=0.000,33.600,49.450,0.0000,0.0000,-110.0000
C00601=150.000,33.600,49.450,0.0000,0.0000,-110.0000
C00602=150.000,29.400,49.450,0.0000,0.0000,-110.0000
C00603=0.000,29.400,49.450,0.0000,0.0000,-110.0000
C00604=0.000,25.200,49.450,0.0000,0.0000,-110.0000
C00605=150.000,25.200,49.450,0.0000,0.0000,-110.0000
C00606=150.000,21.000,49.450,0.0000,0.0000,-110.0000
C00607=0.000,21.000,49.450,0.0000,0.0000,-110.0000
C00608=0.000,16.800,49.450,0.0000,0.0000,-110.0000
C00609=150.000,16.800,49.450,0.0000,0.0000,-110.0000
C00610=150.000,12.600,49.450,0.0000,0.0000,-110.0000
C00611=0.000,12.600,49.450,0.0000,0.0000,-110.0000
C00612=0.000,8.400,49.450,0.0000,0.0000,-110.0000
C00613=150.000,8.400,49.450,0.0000,0.0000,-110.0000
C00614=150.000,4.200,49.450,0.0000,0.0000,-110.0000
C00615=0.000,4.200,49.450,0.0000,0.0000,-110.0000
C00616=0.000,4.200,74.450,0.0000,0.0000,-110.0000
C00617=0.000,0.000,51.600,0.0000,0.0000,-110.0000
C00618=150.000,0.000,51.600,0.0000,0.0000,-110.0000
C00619=0.000,46.200,51.600,0.0000,0.0000,-110.0000
C00620=150.000,46.200,51.600,0.0000,0.0000,-110.0000
C00621=150.000,4.200,51.600,0.0000,0.0000,-110.0000
C00622=0.000,4.200,51.600,0.0000,0.0000,-110.0000
C00623=0.000,8.400,51.600,0.0000,0.0000,-110.0000
C00624=150.000,8.400,51.600,0.0000,0.0000,-110.0000
C00625=150.000,12.600,51.600,0.0000,0.0000,-110.0000
C00626=0.000,12.600,51.600,0.0000,0.0000,-110.0000
C00627=0.000,16.800,51.600,0.0000,0.0000,-110.0000
C00628=150.000,16.800,51.600,0.0000,0.0000,-110.0000
C00629=150.000,21.000,51.600,0.0000,0.0000,-110.0000
C00630=0.000,21.000,51.600,0.0000,0.0000,-110.0000
C00631=0.000,25.200,51.600,0.0000,0.0000,-110.0000
C00632=150.000,25.200,51.600,0.0000,0.0000,-110.0000
C00633=150.000,29.400,51.600,0.0000,0.0000,-110.0000
C00634=0.000,29.400,51.600,0.0000,0.0000,-110.0000
C00635=0.000,33.600,51.600,0.0000,0.0000,-110.0000
C00636=150.000,33.600,51.600,0.0000,0.0000,-110.0000
C00637=150.000,37.800,51.600,0.0000,0.0000,-110.0000
C00638=0.000,37.800,51.600,0.0000,0.0000,-110.0000
C00639=0.000,42.000,51.600,0.0000,0.0000,-110.0000
C00640=150.000,42.000,51.600,0.0000,0.0000,-110.0000
C00641=0.000,0.000,51.600,0.0000,0.0000,-110.0000
C00642=150.000,0.000,51.600,0.0000,0.0000,-110.0000
C00643=0.000,46.200,51.600,0.0000,0.0000,-110.0000
C00644=150.000,46.200,51.600,0.0000,0.0000,-110.0000
C00645=150.000,46.200,76.600,0.0000,0.0000,-110.0000
C00646=150.000,46.200,53.750,0.0000,0.0000,-110.0000
C00647=0.000,46.200,53.750,0.0000,0.0000,-110.0000
C00648=150.000,0.000,53.750,0.0000,0.0000,-110.0000
C00649=0.000,0.000,53.750,0.0000,0.0000,-110.0000
C00650=0.000,42.000,53.750,0.0000,0.0000,-110.0000
C00651=150.000,42.000,53.750,0.0000,0.0000,-110.0000
C00652=150.000,37.800,53.750,0.0000,0.0000,-110.0000
C00653=0.000,37.800,53.750,0.0000,0.0000,-110.0000
C00654=0.000,33.600,53.750,0.0000,0.0000,-110.0000
C00655=150.000,33.600,53.750,0.0000,0.0000,-110.0000
C00656=150.000,29.400,53.750,0.0000,0.0000,-110.0000
C00657=0.000,29.400,53.750,0.0000,0.0000,-110.0000
C00658=0.000,25.200,53.750,0.0000,0.0000,-110.0000
C00659=150.000,25.200,53.750,0.0000,0.0000,-110.0000
C00660=150.000,21.000,53.750,0.0000,0.0000,-110.0000
C00661=0.000,21.000,53.750,0.0000,0.0000,-110.0000
C00662=0.000,16.800,53.750,0.0000,0.0000,-110.0000
C00663=150.000,16.800,53.750,0.0000,0.0000,-110.0000
C00664=150.000,12.600,53.750,0.0000,0.0000,-110.0000
C00665=0.000,12.600,53.750,0.0000,0.0000,-110.0000
C00666=0.000,8.400,53.750,0.0000,0.0000,-110.0000
C00667=150.000,8.400,53.750,0.0000,0.0000,-110.0000
C00668=150.000,4.200,53.750,0.0000,0.0000,-110.0000
C00669=0.000,4.200,53.750,0.0000,0.0000,-110.0000
C00670=0.000,4.200,78.750,0.0000,0.0000,-110.0000
C00671=0.000,0.000,55.900,0.0000,0.0000,-110.0000
C00672=150.000,0.000,55.900,0.0000,0.0000,-110.0000
C00673=0.000,46.200,55.900,0.0000,0.0000,-110.0000
C00674=150.000,46.200,55.900,0.0000,0.0000,-110.0000
C00675=150.000,4.200,55.900,0.0000,0.0000,-110.0000
C00676=0.000,4.200,55.900,0.0000,0.0000,-110.0000
C00677=0.000,8.400,55.900,0.0000,0.0000,-110.0000
C00678=150.000,8.400,55.900,0.0000,0.0000,-110.0000
C00679=150.000,12.600,55.900,0.0000,0.0000,-110.0000
C00680=0.000,12.600,55.900,0.0000,0.0000,-110.0000
C00681=0.000,16.800,55.900,0.0000,0.0000,-110.0000
C00682=150.000,16.800,55.900,0.0000,0.0000,-110.0000
C00683=150.000,21.000,55.900,0.0000,0.0000,-110.0000
C00684=0.000,21.000,55.900,0.0000,0.0000,-110.0000
C00685=0.000,25.200,55.900,0.0000,0.0000,-110.0000
C00686=150.000,25.200,55.900,0.0000,0.0000,-110.0000
C00687=150.000,29.400,55.900,0.0000,0.0000,-110.0000
C00688=0.000,29.400,55.900,0.0000,0.0000,-110.0000
C00689=0.000,33.600,55.900,0.0000,0.0000,-110.0000
C00690=150.000,33.600,55.900,0.0000,0.0000,-110.0000
C00691=150.000,37.800,55.900,0.0000,0.0000,-110.0000
C00692=0.000,37.800,55.900,0.0000,0.0000,-110.0000
C00693=0.000,42.000,55.900,0.0000,0.0000,-110.0000
C00694=150.000,42.000,55.900,0.0000,0.0000,-110.0000
C00695=150.000,42.000,80.900,0.0000,0.0000,-110.0000
C00696=150.000,46.200,58.050,0.0000,0.0000,-110.0000
C00697=0.000,46.200,58.050,0.0000,0.0000,-110.0000
C00698=150.000,0.000,58.050,0.0000,0.0000,-110.0000
C00699=0.000,0.000,58.050,0.0000,0.0000,-110.0000
C00700=0.000,42.000,58.050,0.0000,0.0000,-110.0000
C00701=150.000,42.000,58.050,0.0000,0.0000,-110.0000
C00702=150.000,37.800,58.050,0.0000,0.0000,-110.0000
C00703=0.000,37.800,58.050,0.0000,0.0000,-110.0000
C00704=0.000,33.600,58.050,0.0000,0.0000,-110.0000
C00705=150.000,33.600,58.050,0.0000,0.0000,-110.0000
C00706=150.000,29.400,58.050,0.0000,0.0000,-110.0000
C00707=0.000,29.400,58.050,0.0000,0.0000,-110.0000
C00708=0.000,25.200,58.050,0.0000,0.0000,-110.0000
C00709=150.000,25.200,58.050,0.0000,0.0000,-110.0000
C00710=150.000,21.000,58.050,0.0000,0.0000,-110.0000
C00711=0.000,21.000,58.050,0.0000,0.0000,-110.0000
C00712=0.000,16.800,58.050,0.0000,0.0000,-110.0000
C00713=150.000,16.800,58.050,0.0000,0.0000,-110.0000
C00714=150.000,12.600,58.050,0.0000,0.0000,-110.0000
C00715=0.000,12.600,58.050,0.0000,0.0000,-110.0000
C00716=0.000,8.400,58.050,0.0000,0.0000,-110.0000
C00717=150.000,8.400,58.050,0.0000,0.0000,-110.0000
C00718=150.000,4.200,58.050,0.0000,0.0000,-110.0000
C00719=0.000,4.200,58.050,0.0000,0.0000,-110.0000
C00720=0.000,4.200,83.050,0.0000,0.0000,-110.0000
C00721=0.000,0.000,60.200,0.0000,0.0000,-110.0000
C00722=150.000,0.000,60.200,0.0000,0.0000,-110.0000
C00723=0.000,46.200,60.200,0.0000,0.0000,-110.0000
C00724=150.000,46.200,60.200,0.0000,0.0000,-110.0000
C00725=150.000,4.200,60.200,0.0000,0.0000,-110.0000
C00726=0.000,4.200,60.200,0.0000,0.0000,-110.0000
C00727=0.000,8.400,60.200,0.0000,0.0000,-110.0000
C00728=150.000,8.400,60.200,0.0000,0.0000,-110.0000
C00729=150.000,12.600,60.200,0.0000,0.0000,-110.0000
C00730=0.000,12.600,60.200,0.0000,0.0000,-110.0000
C00731=0.000,16.800,60.200,0.0000,0.0000,-110.0000
C00732=150.000,16.800,60.200,0.0000,0.0000,-110.0000
C00733=150.000,21.000,60.200,0.0000,0.0000,-110.0000
C00734=0.000,21.000,60.200,0.0000,0.0000,-110.0000
C00735=0.000,25.200,60.200,0.0000,0.0000,-110.0000
C00736=150.000,25.200,60.200,0.0000,0.0000,-110.0000
C00737=150.000,29.400,60.200,0.0000,0.0000,-110.0000
C00738=0.000,29.400,60.200,0.0000,0.0000,-110.0000
C00739=0.000,33.600,60.200,0.0000,0.0000,-110.0000
C00740=150.000,33.600,60.200,0.0000,0.0000,-110.0000
C00741=150.000,37.800,60.200,0.0000,0.0000,-110.0000
C00742=0.000,37.800,60.200,0.0000,0.0000,-110.0000
C00743=0.000,42.000,60.200,0.0000,0.0000,-110.0000
C00744=150.000,42.000,60.200,0.0000,0.0000,-110.0000
C00745=150.000,42.000,85.200,0.0000,0.0000,-110.0000
C00746=150.000,46.200,62.350,0.0000,0.0000,-110.0000
C00747=0.000,46.200,62.350,0.0000,0.0000,-110.0000
C00748=150.000,0.000,62.350,0.0000,0.0000,-110.0000
C00749=0.000,0.000,62.350,0.0000,0.0000,-110.0000
C00750=0.000,42.000,62.350,0.0000,0.0000,-110.0000
C00751=150.000,42.000,62.350,0.0000,0.0000,-110.0000
C00752=150.000,37.800,62.350,0.0000,0.0000,-110.0000
C00753=0.000,37.800,62.350,0.0000,0.0000,-110.0000
C00754=0.000,33.600,62.350,0.0000,0.0000,-110.0000
C00755=150.000,33.600,62.350,0.0000,0.0000,-110.0000
C00756=150.000,29.400,62.350,0.0000,0.0000,-110.0000
C00757=0.000,29.400,62.350,0.0000,0.0000,-110.0000
C00758=0.000,25.200,62.350,0.0000,0.0000,-110.0000
C00759=150.000,25.200,62.350,0.0000,0.0000,-110.0000
C00760=150.000,21.000,62.350,0.0000,0.0000,-110.0000
C00761=0.000,21.000,62.350,0.0000,0.0000,-110.0000
C00762=0.000,16.800,62.350,0.0000,0.0000,-110.0000
C00763=150.000,16.800,62.350,0.0000,0.0000,-110.0000
C00764=150.000,12.600,62.350,0.0000,0.0000,-110.0000
C00765=0.000,12.600,62.350,0.0000,0.0000,-110.0000
C00766=0.000,8.400,62.350,0.0000,0.0000,-110.0000
C00767=150.000,8.400,62.350,0.0000,0.0000,-110.0000
C00768=150.000,4.200,62.350,0.0000,0.0000,-110.0000
C00769=0.000,4.200,62.350,0.0000,0.0000,-110.0000
C00770=150.000,46.200,62.350,0.0000,0.0000,-110.0000
C00771=0.000,46.200,62.350,0.0000,0.0000,-110.0000
C00772=150.000,0.000,62.350,0.0000,0.0000,-110.0000
C00773=0.000,0.000,62.350,0.0000,0.0000,-110.0000
C00774=0.000,0.000,87.350,0.0000,0.0000,-110.0000
//INST
///DATE 2026/09/11 12:21
///COMM Python Generated
///ATTR SC,RW,RJ
////FRAME USER 3
///GROUP1 RB1
NOP
DOUT OT#(9) OFF
TIMER T=5.00
MOVJ C00000 VJ=10.00 ACC=20
*LABEL0
MOVJ C00001 VJ=10.00 ACC=20
MACRO1 MJ#(0) ARGF103
ARCON
MOVL C00002 V=13.5 ACC=20
ARCOF
TIMER T=7.00
*LABEL1
MOVJ C00003 VJ=10.00 ACC=20
MACRO1 MJ#(0) ARGF103
ARCON
MOVL C00004 V=13.5 ACC=20
ARCOF
TIMER T=7.00
*LABEL2
MOVJ C00005 VJ=10.00 ACC=20
MACRO1 MJ#(0) ARGF101
ARCON
MOVL C00006 V=13.5 ACC=20
ARCOF
TIMER T=7.00
*LABEL3
MOVJ C00007 VJ=10.00 ACC=20
MACRO1 MJ#(0) ARGF101
ARCON
MOVL C00008 V=13.5 ACC=20
ARCOF
TIMER T=7.00
*LABEL4
MOVJ C00009 VJ=10.00 ACC=20
MACRO1 MJ#(0) ARGF101
ARCON
MOVL C00010 V=13.5 ACC=20
ARCOF
TIMER T=7.00
*LABEL5
MOVJ C00011 VJ=10.00 ACC=20
MACRO1 MJ#(0) ARGF101
ARCON
MOVL C00012 V=13.5 ACC=20
ARCOF
TIMER T=7.00
*LABEL6
MOVJ C00013 VJ=10.00 ACC=20
MACRO1 MJ#(0) ARGF101
ARCON
MOVL C00014 V=13.5 ACC=20
ARCOF
TIMER T=7.00
*LABEL7
MOVJ C00015 VJ=10.00 ACC=20
MACRO1 MJ#(0) ARGF101
ARCON
MOVL C00016 V=13.5 ACC=20
ARCOF
TIMER T=7.00
*LABEL8
MOVJ C00017 VJ=10.00 ACC=20
MACRO1 MJ#(0) ARGF101
ARCON
MOVL C00018 V=13.5 ACC=20
ARCOF
TIMER T=7.00
*LABEL9
MOVJ C00019 VJ=10.00 ACC=20
MACRO1 MJ#(0) ARGF101
ARCON
MOVL C00020 V=13.5 ACC=20
ARCOF
TIMER T=7.00
*LABEL10
MOVJ C00021 VJ=10.00 ACC=20
MACRO1 MJ#(0) ARGF101
ARCON
MOVL C00022 V=13.5 ACC=20
ARCOF
TIMER T=7.00
*LABEL11
MOVJ C00023 VJ=10.00 ACC=20
MACRO1 MJ#(0) ARGF101
ARCON
MOVL C00024 V=13.5 ACC=20
ARCOF
DOUT OT#(9) ON
TIMER T=50.00
DOUT OT#(9) OFF
TIMER T=13.00
MOVJ C00025 VJ=10.00 ACC=20
*LABEL12
MOVJ C00026 VJ=10.00 ACC=20
MACRO1 MJ#(0) ARGF103
ARCON
MOVL C00027 V=13.5 ACC=20
ARCOF
TIMER T=7.00
*LABEL13
MOVJ C00028 VJ=10.00 ACC=20
MACRO1 MJ#(0) ARGF103
ARCON
MOVL C00029 V=13.5 ACC=20
ARCOF
TIMER T=7.00
*LABEL14
MOVJ C00030 VJ=10.00 ACC=20
MACRO1 MJ#(0) ARGF101
ARCON
MOVL C00031 V=13.5 ACC=20
ARCOF
TIMER T=7.00
*LABEL15
MOVJ C00032 VJ=10.00 ACC=20
MACRO1 MJ#(0) ARGF101
ARCON
MOVL C00033 V=13.5 ACC=20
ARCOF
TIMER T=7.00
*LABEL16
MOVJ C00034 VJ=10.00 ACC=20
MACRO1 MJ#(0) ARGF101
ARCON
MOVL C00035 V=13.5 ACC=20
ARCOF
TIMER T=7.00
*LABEL17
MOVJ C00036 VJ=10.00 ACC=20
MACRO1 MJ#(0) ARGF101
ARCON
MOVL C00037 V=13.5 ACC=20
ARCOF
TIMER T=7.00
*LABEL18
MOVJ C00038 VJ=10.00 ACC=20
MACRO1 MJ#(0) ARGF101
ARCON
MOVL C00039 V=13.5 ACC=20
ARCOF
TIMER T=7.00
*LABEL19
MOVJ C00040 VJ=10.00 ACC=20
MACRO1 MJ#(0) ARGF101
ARCON
MOVL C00041 V=13.5 ACC=20
ARCOF
TIMER T=7.00
*LABEL20
MOVJ C00042 VJ=10.00 ACC=20
MACRO1 MJ#(0) ARGF101
ARCON
MOVL C00043 V=13.5 ACC=20
ARCOF
TIMER T=7.00
*LABEL21
MOVJ C00044 VJ=10.00 ACC=20
MACRO1 MJ#(0) ARGF101
ARCON
MOVL C00045 V=13.5 ACC=20
ARCOF
TIMER T=7.00
*LABEL22
MOVJ C00046 VJ=10.00 ACC=20
MACRO1 MJ#(0) ARGF101
ARCON
MOVL C00047 V=13.5 ACC=20
ARCOF
TIMER T=7.00
*LABEL23
MOVJ C00048 VJ=10.00 ACC=20
MACRO1 MJ#(0) ARGF101
ARCON
MOVL C00049 V=13.5 ACC=20
ARCOF
DOUT OT#(9) ON
TIMER T=50.00
DOUT OT#(9) OFF
TIMER T=13.00
MOVJ C00050 VJ=10.00 ACC=20
*LABEL24
MOVJ C00051 VJ=10.00 ACC=20
MACRO1 MJ#(0) ARGF103
ARCON
MOVL C00052 V=13.5 ACC=20
ARCOF
TIMER T=7.00
*LABEL25
MOVJ C00053 VJ=10.00 ACC=20
MACRO1 MJ#(0) ARGF103
ARCON
MOVL C00054 V=13.5 ACC=20
ARCOF
TIMER T=7.00
*LABEL26
MOVJ C00055 VJ=10.00 ACC=20
MACRO1 MJ#(0) ARGF101
ARCON
MOVL C00056 V=13.5 ACC=20
ARCOF
TIMER T=7.00
*LABEL27
MOVJ C00057 VJ=10.00 ACC=20
MACRO1 MJ#(0) ARGF101
ARCON
MOVL C00058 V=13.5 ACC=20
ARCOF
TIMER T=7.00
*LABEL28
MOVJ C00059 VJ=10.00 ACC=20
MACRO1 MJ#(0) ARGF101
ARCON
MOVL C00060 V=13.5 ACC=20
ARCOF
TIMER T=7.00
*LABEL29
MOVJ C00061 VJ=10.00 ACC=20
MACRO1 MJ#(0) ARGF101
ARCON
MOVL C00062 V=13.5 ACC=20
ARCOF
TIMER T=7.00
*LABEL30
MOVJ C00063 VJ=10.00 ACC=20
MACRO1 MJ#(0) ARGF101
ARCON
MOVL C00064 V=13.5 ACC=20
ARCOF
TIMER T=7.00
*LABEL31
MOVJ C00065 VJ=10.00 ACC=20
MACRO1 MJ#(0) ARGF101
ARCON
MOVL C00066 V=13.5 ACC=20
ARCOF
TIMER T=7.00
*LABEL32
MOVJ C00067 VJ=10.00 ACC=20
MACRO1 MJ#(0) ARGF101
ARCON
MOVL C00068 V=13.5 ACC=20
ARCOF
TIMER T=7.00
*LABEL33
MOVJ C00069 VJ=10.00 ACC=20
MACRO1 MJ#(0) ARGF101
ARCON
MOVL C00070 V=13.5 ACC=20
ARCOF
TIMER T=7.00
*LABEL34
MOVJ C00071 VJ=10.00 ACC=20
MACRO1 MJ#(0) ARGF101
ARCON
MOVL C00072 V=13.5 ACC=20
ARCOF
TIMER T=7.00
*LABEL35
MOVJ C00073 VJ=10.00 ACC=20
MACRO1 MJ#(0) ARGF101
ARCON
MOVL C00074 V=13.5 ACC=20
ARCOF
DOUT OT#(9) ON
TIMER T=50.00
DOUT OT#(9) OFF
TIMER T=13.00
MOVJ C00075 VJ=10.00 ACC=20
*LABEL36
MOVJ C00076 VJ=10.00 ACC=20
MACRO1 MJ#(0) ARGF103
ARCON
MOVL C00077 V=13.5 ACC=20
ARCOF
TIMER T=7.00
*LABEL37
MOVJ C00078 VJ=10.00 ACC=20
MACRO1 MJ#(0) ARGF103
ARCON
MOVL C00079 V=13.5 ACC=20
ARCOF
TIMER T=7.00
*LABEL38
MOVJ C00080 VJ=10.00 ACC=20
MACRO1 MJ#(0) ARGF101
ARCON
MOVL C00081 V=13.5 ACC=20
ARCOF
TIMER T=7.00
*LABEL39
MOVJ C00082 VJ=10.00 ACC=20
MACRO1 MJ#(0) ARGF101
ARCON
MOVL C00083 V=13.5 ACC=20
ARCOF
TIMER T=7.00
*LABEL40
MOVJ C00084 VJ=10.00 ACC=20
MACRO1 MJ#(0) ARGF101
ARCON
MOVL C00085 V=13.5 ACC=20
ARCOF
TIMER T=7.00
*LABEL41
MOVJ C00086 VJ=10.00 ACC=20
MACRO1 MJ#(0) ARGF101
ARCON
MOVL C00087 V=13.5 ACC=20
ARCOF
TIMER T=7.00
*LABEL42
MOVJ C00088 VJ=10.00 ACC=20
MACRO1 MJ#(0) ARGF101
ARCON
MOVL C00089 V=13.5 ACC=20
ARCOF
TIMER T=7.00
*LABEL43
MOVJ C00090 VJ=10.00 ACC=20
MACRO1 MJ#(0) ARGF101
ARCON
MOVL C00091 V=13.5 ACC=20
ARCOF
TIMER T=7.00
*LABEL44
MOVJ C00092 VJ=10.00 ACC=20
MACRO1 MJ#(0) ARGF101
ARCON
MOVL C00093 V=13.5 ACC=20
ARCOF
TIMER T=7.00
*LABEL45
MOVJ C00094 VJ=10.00 ACC=20
MACRO1 MJ#(0) ARGF101
ARCON
MOVL C00095 V=13.5 ACC=20
ARCOF
TIMER T=7.00
*LABEL46
MOVJ C00096 VJ=10.00 ACC=20
MACRO1 MJ#(0) ARGF101
ARCON
MOVL C00097 V=13.5 ACC=20
ARCOF
TIMER T=7.00
*LABEL47
MOVJ C00098 VJ=10.00 ACC=20
MACRO1 MJ#(0) ARGF101
ARCON
MOVL C00099 V=13.5 ACC=20
ARCOF
DOUT OT#(9) ON
TIMER T=50.00
DOUT OT#(9) OFF
TIMER T=13.00
MOVJ C00100 VJ=10.00 ACC=20
*LABEL48
MOVJ C00101 VJ=10.00 ACC=20
MACRO1 MJ#(0) ARGF103
ARCON
MOVL C00102 V=13.5 ACC=20
ARCOF
TIMER T=7.00
*LABEL49
MOVJ C00103 VJ=10.00 ACC=20
MACRO1 MJ#(0) ARGF103
ARCON
MOVL C00104 V=13.5 ACC=20
ARCOF
TIMER T=7.00
*LABEL50
MOVJ C00105 VJ=10.00 ACC=20
MACRO1 MJ#(0) ARGF101
ARCON
MOVL C00106 V=13.5 ACC=20
ARCOF
TIMER T=7.00
*LABEL51
MOVJ C00107 VJ=10.00 ACC=20
MACRO1 MJ#(0) ARGF101
ARCON
MOVL C00108 V=13.5 ACC=20
ARCOF
TIMER T=7.00
*LABEL52
MOVJ C00109 VJ=10.00 ACC=20
MACRO1 MJ#(0) ARGF101
ARCON
MOVL C00110 V=13.5 ACC=20
ARCOF
TIMER T=7.00
*LABEL53
MOVJ C00111 VJ=10.00 ACC=20
MACRO1 MJ#(0) ARGF101
ARCON
MOVL C00112 V=13.5 ACC=20
ARCOF
TIMER T=7.00
*LABEL54
MOVJ C00113 VJ=10.00 ACC=20
MACRO1 MJ#(0) ARGF101
ARCON
MOVL C00114 V=13.5 ACC=20
ARCOF
TIMER T=7.00
*LABEL55
MOVJ C00115 VJ=10.00 ACC=20
MACRO1 MJ#(0) ARGF101
ARCON
MOVL C00116 V=13.5 ACC=20
ARCOF
TIMER T=7.00
*LABEL56
MOVJ C00117 VJ=10.00 ACC=20
MACRO1 MJ#(0) ARGF101
ARCON
MOVL C00118 V=13.5 ACC=20
ARCOF
TIMER T=7.00
*LABEL57
MOVJ C00119 VJ=10.00 ACC=20
MACRO1 MJ#(0) ARGF101
ARCON
MOVL C00120 V=13.5 ACC=20
ARCOF
TIMER T=7.00
*LABEL58
MOVJ C00121 VJ=10.00 ACC=20
MACRO1 MJ#(0) ARGF101
ARCON
MOVL C00122 V=13.5 ACC=20
ARCOF
TIMER T=7.00
*LABEL59
MOVJ C00123 VJ=10.00 ACC=20
MACRO1 MJ#(0) ARGF101
ARCON
MOVL C00124 V=13.5 ACC=20
ARCOF
TIMER T=7.00
*LABEL60
MOVJ C00125 VJ=10.00 ACC=20
MACRO1 MJ#(0) ARGF103
ARCON
MOVL C00126 V=13.5 ACC=20
ARCOF
TIMER T=7.00
*LABEL61
MOVJ C00127 VJ=10.00 ACC=20
MACRO1 MJ#(0) ARGF103
ARCON
MOVL C00128 V=13.5 ACC=20
ARCOF
DOUT OT#(9) ON
TIMER T=50.00
DOUT OT#(9) OFF
TIMER T=13.00
MOVJ C00129 VJ=10.00 ACC=20
*LABEL62
MOVJ C00130 VJ=10.00 ACC=20
MACRO1 MJ#(0) ARGF103
ARCON
MOVL C00131 V=13.5 ACC=20
ARCOF
TIMER T=7.00
*LABEL63
MOVJ C00132 VJ=10.00 ACC=20
MACRO1 MJ#(0) ARGF103
ARCON
MOVL C00133 V=13.5 ACC=20
ARCOF
TIMER T=7.00
*LABEL64
MOVJ C00134 VJ=10.00 ACC=20
MACRO1 MJ#(0) ARGF101
ARCON
MOVL C00135 V=13.5 ACC=20
ARCOF
TIMER T=7.00
*LABEL65
MOVJ C00136 VJ=10.00 ACC=20
MACRO1 MJ#(0) ARGF101
ARCON
MOVL C00137 V=13.5 ACC=20
ARCOF
TIMER T=7.00
*LABEL66
MOVJ C00138 VJ=10.00 ACC=20
MACRO1 MJ#(0) ARGF101
ARCON
MOVL C00139 V=13.5 ACC=20
ARCOF
TIMER T=7.00
*LABEL67
MOVJ C00140 VJ=10.00 ACC=20
MACRO1 MJ#(0) ARGF101
ARCON
MOVL C00141 V=13.5 ACC=20
ARCOF
TIMER T=7.00
*LABEL68
MOVJ C00142 VJ=10.00 ACC=20
MACRO1 MJ#(0) ARGF101
ARCON
MOVL C00143 V=13.5 ACC=20
ARCOF
TIMER T=7.00
*LABEL69
MOVJ C00144 VJ=10.00 ACC=20
MACRO1 MJ#(0) ARGF101
ARCON
MOVL C00145 V=13.5 ACC=20
ARCOF
TIMER T=7.00
*LABEL70
MOVJ C00146 VJ=10.00 ACC=20
MACRO1 MJ#(0) ARGF101
ARCON
MOVL C00147 V=13.5 ACC=20
ARCOF
TIMER T=7.00
*LABEL71
MOVJ C00148 VJ=10.00 ACC=20
MACRO1 MJ#(0) ARGF101
ARCON
MOVL C00149 V=13.5 ACC=20
ARCOF
TIMER T=7.00
*LABEL72
MOVJ C00150 VJ=10.00 ACC=20
MACRO1 MJ#(0) ARGF101
ARCON
MOVL C00151 V=13.5 ACC=20
ARCOF
TIMER T=7.00
*LABEL73
MOVJ C00152 VJ=10.00 ACC=20
MACRO1 MJ#(0) ARGF101
ARCON
MOVL C00153 V=13.5 ACC=20
ARCOF
DOUT OT#(9) ON
TIMER T=50.00
DOUT OT#(9) OFF
TIMER T=13.00
MOVJ C00154 VJ=10.00 ACC=20
*LABEL74
MOVJ C00155 VJ=10.00 ACC=20
MACRO1 MJ#(0) ARGF103
ARCON
MOVL C00156 V=13.5 ACC=20
ARCOF
TIMER T=7.00
*LABEL75
MOVJ C00157 VJ=10.00 ACC=20
MACRO1 MJ#(0) ARGF103
ARCON
MOVL C00158 V=13.5 ACC=20
ARCOF
TIMER T=7.00
*LABEL76
MOVJ C00159 VJ=10.00 ACC=20
MACRO1 MJ#(0) ARGF101
ARCON
MOVL C00160 V=13.5 ACC=20
ARCOF
TIMER T=7.00
*LABEL77
MOVJ C00161 VJ=10.00 ACC=20
MACRO1 MJ#(0) ARGF101
ARCON
MOVL C00162 V=13.5 ACC=20
ARCOF
TIMER T=7.00
*LABEL78
MOVJ C00163 VJ=10.00 ACC=20
MACRO1 MJ#(0) ARGF101
ARCON
MOVL C00164 V=13.5 ACC=20
ARCOF
TIMER T=7.00
*LABEL79
MOVJ C00165 VJ=10.00 ACC=20
MACRO1 MJ#(0) ARGF101
ARCON
MOVL C00166 V=13.5 ACC=20
ARCOF
TIMER T=7.00
*LABEL80
MOVJ C00167 VJ=10.00 ACC=20
MACRO1 MJ#(0) ARGF101
ARCON
MOVL C00168 V=13.5 ACC=20
ARCOF
TIMER T=7.00
*LABEL81
MOVJ C00169 VJ=10.00 ACC=20
MACRO1 MJ#(0) ARGF101
ARCON
MOVL C00170 V=13.5 ACC=20
ARCOF
TIMER T=7.00
*LABEL82
MOVJ C00171 VJ=10.00 ACC=20
MACRO1 MJ#(0) ARGF101
ARCON
MOVL C00172 V=13.5 ACC=20
ARCOF
TIMER T=7.00
*LABEL83
MOVJ C00173 VJ=10.00 ACC=20
MACRO1 MJ#(0) ARGF101
ARCON
MOVL C00174 V=13.5 ACC=20
ARCOF
TIMER T=7.00
*LABEL84
MOVJ C00175 VJ=10.00 ACC=20
MACRO1 MJ#(0) ARGF101
ARCON
MOVL C00176 V=13.5 ACC=20
ARCOF
TIMER T=7.00
*LABEL85
MOVJ C00177 VJ=10.00 ACC=20
MACRO1 MJ#(0) ARGF101
ARCON
MOVL C00178 V=13.5 ACC=20
ARCOF
DOUT OT#(9) ON
TIMER T=50.00
DOUT OT#(9) OFF
TIMER T=13.00
MOVJ C00179 VJ=10.00 ACC=20
*LABEL86
MOVJ C00180 VJ=10.00 ACC=20
MACRO1 MJ#(0) ARGF103
ARCON
MOVL C00181 V=13.5 ACC=20
ARCOF
TIMER T=7.00
*LABEL87
MOVJ C00182 VJ=10.00 ACC=20
MACRO1 MJ#(0) ARGF103
ARCON
MOVL C00183 V=13.5 ACC=20
ARCOF
TIMER T=7.00
*LABEL88
MOVJ C00184 VJ=10.00 ACC=20
MACRO1 MJ#(0) ARGF101
ARCON
MOVL C00185 V=13.5 ACC=20
ARCOF
TIMER T=7.00
*LABEL89
MOVJ C00186 VJ=10.00 ACC=20
MACRO1 MJ#(0) ARGF101
ARCON
MOVL C00187 V=13.5 ACC=20
ARCOF
TIMER T=7.00
*LABEL90
MOVJ C00188 VJ=10.00 ACC=20
MACRO1 MJ#(0) ARGF101
ARCON
MOVL C00189 V=13.5 ACC=20
ARCOF
TIMER T=7.00
*LABEL91
MOVJ C00190 VJ=10.00 ACC=20
MACRO1 MJ#(0) ARGF101
ARCON
MOVL C00191 V=13.5 ACC=20
ARCOF
TIMER T=7.00
*LABEL92
MOVJ C00192 VJ=10.00 ACC=20
MACRO1 MJ#(0) ARGF101
ARCON
MOVL C00193 V=13.5 ACC=20
ARCOF
TIMER T=7.00
*LABEL93
MOVJ C00194 VJ=10.00 ACC=20
MACRO1 MJ#(0) ARGF101
ARCON
MOVL C00195 V=13.5 ACC=20
ARCOF
TIMER T=7.00
*LABEL94
MOVJ C00196 VJ=10.00 ACC=20
MACRO1 MJ#(0) ARGF101
ARCON
MOVL C00197 V=13.5 ACC=20
ARCOF
TIMER T=7.00
*LABEL95
MOVJ C00198 VJ=10.00 ACC=20
MACRO1 MJ#(0) ARGF101
ARCON
MOVL C00199 V=13.5 ACC=20
ARCOF
TIMER T=7.00
*LABEL96
MOVJ C00200 VJ=10.00 ACC=20
MACRO1 MJ#(0) ARGF101
ARCON
MOVL C00201 V=13.5 ACC=20
ARCOF
TIMER T=7.00
*LABEL97
MOVJ C00202 VJ=10.00 ACC=20
MACRO1 MJ#(0) ARGF101
ARCON
MOVL C00203 V=13.5 ACC=20
ARCOF
DOUT OT#(9) ON
TIMER T=50.00
DOUT OT#(9) OFF
TIMER T=13.00
MOVJ C00204 VJ=10.00 ACC=20
*LABEL98
MOVJ C00205 VJ=10.00 ACC=20
MACRO1 MJ#(0) ARGF103
ARCON
MOVL C00206 V=13.5 ACC=20
ARCOF
TIMER T=7.00
*LABEL99
MOVJ C00207 VJ=10.00 ACC=20
MACRO1 MJ#(0) ARGF103
ARCON
MOVL C00208 V=13.5 ACC=20
ARCOF
TIMER T=7.00
*LABEL100
MOVJ C00209 VJ=10.00 ACC=20
MACRO1 MJ#(0) ARGF101
ARCON
MOVL C00210 V=13.5 ACC=20
ARCOF
TIMER T=7.00
*LABEL101
MOVJ C00211 VJ=10.00 ACC=20
MACRO1 MJ#(0) ARGF101
ARCON
MOVL C00212 V=13.5 ACC=20
ARCOF
TIMER T=7.00
*LABEL102
MOVJ C00213 VJ=10.00 ACC=20
MACRO1 MJ#(0) ARGF101
ARCON
MOVL C00214 V=13.5 ACC=20
ARCOF
TIMER T=7.00
*LABEL103
MOVJ C00215 VJ=10.00 ACC=20
MACRO1 MJ#(0) ARGF101
ARCON
MOVL C00216 V=13.5 ACC=20
ARCOF
TIMER T=7.00
*LABEL104
MOVJ C00217 VJ=10.00 ACC=20
MACRO1 MJ#(0) ARGF101
ARCON
MOVL C00218 V=13.5 ACC=20
ARCOF
TIMER T=7.00
*LABEL105
MOVJ C00219 VJ=10.00 ACC=20
MACRO1 MJ#(0) ARGF101
ARCON
MOVL C00220 V=13.5 ACC=20
ARCOF
TIMER T=7.00
*LABEL106
MOVJ C00221 VJ=10.00 ACC=20
MACRO1 MJ#(0) ARGF101
ARCON
MOVL C00222 V=13.5 ACC=20
ARCOF
TIMER T=7.00
*LABEL107
MOVJ C00223 VJ=10.00 ACC=20
MACRO1 MJ#(0) ARGF101
ARCON
MOVL C00224 V=13.5 ACC=20
ARCOF
TIMER T=7.00
*LABEL108
MOVJ C00225 VJ=10.00 ACC=20
MACRO1 MJ#(0) ARGF101
ARCON
MOVL C00226 V=13.5 ACC=20
ARCOF
TIMER T=7.00
*LABEL109
MOVJ C00227 VJ=10.00 ACC=20
MACRO1 MJ#(0) ARGF101
ARCON
MOVL C00228 V=13.5 ACC=20
ARCOF
DOUT OT#(9) ON
TIMER T=50.00
DOUT OT#(9) OFF
TIMER T=13.00
MOVJ C00229 VJ=10.00 ACC=20
*LABEL110
MOVJ C00230 VJ=10.00 ACC=20
MACRO1 MJ#(0) ARGF103
ARCON
MOVL C00231 V=13.5 ACC=20
ARCOF
TIMER T=7.00
*LABEL111
MOVJ C00232 VJ=10.00 ACC=20
MACRO1 MJ#(0) ARGF103
ARCON
MOVL C00233 V=13.5 ACC=20
ARCOF
TIMER T=7.00
*LABEL112
MOVJ C00234 VJ=10.00 ACC=20
MACRO1 MJ#(0) ARGF101
ARCON
MOVL C00235 V=13.5 ACC=20
ARCOF
TIMER T=7.00
*LABEL113
MOVJ C00236 VJ=10.00 ACC=20
MACRO1 MJ#(0) ARGF101
ARCON
MOVL C00237 V=13.5 ACC=20
ARCOF
TIMER T=7.00
*LABEL114
MOVJ C00238 VJ=10.00 ACC=20
MACRO1 MJ#(0) ARGF101
ARCON
MOVL C00239 V=13.5 ACC=20
ARCOF
TIMER T=7.00
*LABEL115
MOVJ C00240 VJ=10.00 ACC=20
MACRO1 MJ#(0) ARGF101
ARCON
MOVL C00241 V=13.5 ACC=20
ARCOF
TIMER T=7.00
*LABEL116
MOVJ C00242 VJ=10.00 ACC=20
MACRO1 MJ#(0) ARGF101
ARCON
MOVL C00243 V=13.5 ACC=20
ARCOF
TIMER T=7.00
*LABEL117
MOVJ C00244 VJ=10.00 ACC=20
MACRO1 MJ#(0) ARGF101
ARCON
MOVL C00245 V=13.5 ACC=20
ARCOF
TIMER T=7.00
*LABEL118
MOVJ C00246 VJ=10.00 ACC=20
MACRO1 MJ#(0) ARGF101
ARCON
MOVL C00247 V=13.5 ACC=20
ARCOF
TIMER T=7.00
*LABEL119
MOVJ C00248 VJ=10.00 ACC=20
MACRO1 MJ#(0) ARGF101
ARCON
MOVL C00249 V=13.5 ACC=20
ARCOF
TIMER T=7.00
*LABEL120
MOVJ C00250 VJ=10.00 ACC=20
MACRO1 MJ#(0) ARGF101
ARCON
MOVL C00251 V=13.5 ACC=20
ARCOF
TIMER T=7.00
*LABEL121
MOVJ C00252 VJ=10.00 ACC=20
MACRO1 MJ#(0) ARGF101
ARCON
MOVL C00253 V=13.5 ACC=20
ARCOF
TIMER T=7.00
*LABEL122
MOVJ C00254 VJ=10.00 ACC=20
MACRO1 MJ#(0) ARGF103
ARCON
MOVL C00255 V=13.5 ACC=20
ARCOF
TIMER T=7.00
*LABEL123
MOVJ C00256 VJ=10.00 ACC=20
MACRO1 MJ#(0) ARGF103
ARCON
MOVL C00257 V=13.5 ACC=20
ARCOF
DOUT OT#(9) ON
TIMER T=50.00
DOUT OT#(9) OFF
TIMER T=13.00
MOVJ C00258 VJ=10.00 ACC=20
*LABEL124
MOVJ C00259 VJ=10.00 ACC=20
MACRO1 MJ#(0) ARGF103
ARCON
MOVL C00260 V=13.5 ACC=20
ARCOF
TIMER T=7.00
*LABEL125
MOVJ C00261 VJ=10.00 ACC=20
MACRO1 MJ#(0) ARGF103
ARCON
MOVL C00262 V=13.5 ACC=20
ARCOF
TIMER T=7.00
*LABEL126
MOVJ C00263 VJ=10.00 ACC=20
MACRO1 MJ#(0) ARGF101
ARCON
MOVL C00264 V=13.5 ACC=20
ARCOF
TIMER T=7.00
*LABEL127
MOVJ C00265 VJ=10.00 ACC=20
MACRO1 MJ#(0) ARGF101
ARCON
MOVL C00266 V=13.5 ACC=20
ARCOF
TIMER T=7.00
*LABEL128
MOVJ C00267 VJ=10.00 ACC=20
MACRO1 MJ#(0) ARGF101
ARCON
MOVL C00268 V=13.5 ACC=20
ARCOF
TIMER T=7.00
*LABEL129
MOVJ C00269 VJ=10.00 ACC=20
MACRO1 MJ#(0) ARGF101
ARCON
MOVL C00270 V=13.5 ACC=20
ARCOF
TIMER T=7.00
*LABEL130
MOVJ C00271 VJ=10.00 ACC=20
MACRO1 MJ#(0) ARGF101
ARCON
MOVL C00272 V=13.5 ACC=20
ARCOF
TIMER T=7.00
*LABEL131
MOVJ C00273 VJ=10.00 ACC=20
MACRO1 MJ#(0) ARGF101
ARCON
MOVL C00274 V=13.5 ACC=20
ARCOF
TIMER T=7.00
*LABEL132
MOVJ C00275 VJ=10.00 ACC=20
MACRO1 MJ#(0) ARGF101
ARCON
MOVL C00276 V=13.5 ACC=20
ARCOF
TIMER T=7.00
*LABEL133
MOVJ C00277 VJ=10.00 ACC=20
MACRO1 MJ#(0) ARGF101
ARCON
MOVL C00278 V=13.5 ACC=20
ARCOF
TIMER T=7.00
*LABEL134
MOVJ C00279 VJ=10.00 ACC=20
MACRO1 MJ#(0) ARGF101
ARCON
MOVL C00280 V=13.5 ACC=20
ARCOF
TIMER T=7.00
*LABEL135
MOVJ C00281 VJ=10.00 ACC=20
MACRO1 MJ#(0) ARGF101
ARCON
MOVL C00282 V=13.5 ACC=20
ARCOF
DOUT OT#(9) ON
TIMER T=50.00
DOUT OT#(9) OFF
TIMER T=13.00
MOVJ C00283 VJ=10.00 ACC=20
*LABEL136
MOVJ C00284 VJ=10.00 ACC=20
MACRO1 MJ#(0) ARGF103
ARCON
MOVL C00285 V=13.5 ACC=20
ARCOF
TIMER T=7.00
*LABEL137
MOVJ C00286 VJ=10.00 ACC=20
MACRO1 MJ#(0) ARGF103
ARCON
MOVL C00287 V=13.5 ACC=20
ARCOF
TIMER T=7.00
*LABEL138
MOVJ C00288 VJ=10.00 ACC=20
MACRO1 MJ#(0) ARGF101
ARCON
MOVL C00289 V=13.5 ACC=20
ARCOF
TIMER T=7.00
*LABEL139
MOVJ C00290 VJ=10.00 ACC=20
MACRO1 MJ#(0) ARGF101
ARCON
MOVL C00291 V=13.5 ACC=20
ARCOF
TIMER T=7.00
*LABEL140
MOVJ C00292 VJ=10.00 ACC=20
MACRO1 MJ#(0) ARGF101
ARCON
MOVL C00293 V=13.5 ACC=20
ARCOF
TIMER T=7.00
*LABEL141
MOVJ C00294 VJ=10.00 ACC=20
MACRO1 MJ#(0) ARGF101
ARCON
MOVL C00295 V=13.5 ACC=20
ARCOF
TIMER T=7.00
*LABEL142
MOVJ C00296 VJ=10.00 ACC=20
MACRO1 MJ#(0) ARGF101
ARCON
MOVL C00297 V=13.5 ACC=20
ARCOF
TIMER T=7.00
*LABEL143
MOVJ C00298 VJ=10.00 ACC=20
MACRO1 MJ#(0) ARGF101
ARCON
MOVL C00299 V=13.5 ACC=20
ARCOF
TIMER T=7.00
*LABEL144
MOVJ C00300 VJ=10.00 ACC=20
MACRO1 MJ#(0) ARGF101
ARCON
MOVL C00301 V=13.5 ACC=20
ARCOF
TIMER T=7.00
*LABEL145
MOVJ C00302 VJ=10.00 ACC=20
MACRO1 MJ#(0) ARGF101
ARCON
MOVL C00303 V=13.5 ACC=20
ARCOF
TIMER T=7.00
*LABEL146
MOVJ C00304 VJ=10.00 ACC=20
MACRO1 MJ#(0) ARGF101
ARCON
MOVL C00305 V=13.5 ACC=20
ARCOF
TIMER T=7.00
*LABEL147
MOVJ C00306 VJ=10.00 ACC=20
MACRO1 MJ#(0) ARGF101
ARCON
MOVL C00307 V=13.5 ACC=20
ARCOF
DOUT OT#(9) ON
TIMER T=50.00
DOUT OT#(9) OFF
TIMER T=13.00
MOVJ C00308 VJ=10.00 ACC=20
*LABEL148
MOVJ C00309 VJ=10.00 ACC=20
MACRO1 MJ#(0) ARGF103
ARCON
MOVL C00310 V=13.5 ACC=20
ARCOF
TIMER T=7.00
*LABEL149
MOVJ C00311 VJ=10.00 ACC=20
MACRO1 MJ#(0) ARGF103
ARCON
MOVL C00312 V=13.5 ACC=20
ARCOF
TIMER T=7.00
*LABEL150
MOVJ C00313 VJ=10.00 ACC=20
MACRO1 MJ#(0) ARGF101
ARCON
MOVL C00314 V=13.5 ACC=20
ARCOF
TIMER T=7.00
*LABEL151
MOVJ C00315 VJ=10.00 ACC=20
MACRO1 MJ#(0) ARGF101
ARCON
MOVL C00316 V=13.5 ACC=20
ARCOF
TIMER T=7.00
*LABEL152
MOVJ C00317 VJ=10.00 ACC=20
MACRO1 MJ#(0) ARGF101
ARCON
MOVL C00318 V=13.5 ACC=20
ARCOF
TIMER T=7.00
*LABEL153
MOVJ C00319 VJ=10.00 ACC=20
MACRO1 MJ#(0) ARGF101
ARCON
MOVL C00320 V=13.5 ACC=20
ARCOF
TIMER T=7.00
*LABEL154
MOVJ C00321 VJ=10.00 ACC=20
MACRO1 MJ#(0) ARGF101
ARCON
MOVL C00322 V=13.5 ACC=20
ARCOF
TIMER T=7.00
*LABEL155
MOVJ C00323 VJ=10.00 ACC=20
MACRO1 MJ#(0) ARGF101
ARCON
MOVL C00324 V=13.5 ACC=20
ARCOF
TIMER T=7.00
*LABEL156
MOVJ C00325 VJ=10.00 ACC=20
MACRO1 MJ#(0) ARGF101
ARCON
MOVL C00326 V=13.5 ACC=20
ARCOF
TIMER T=7.00
*LABEL157
MOVJ C00327 VJ=10.00 ACC=20
MACRO1 MJ#(0) ARGF101
ARCON
MOVL C00328 V=13.5 ACC=20
ARCOF
TIMER T=7.00
*LABEL158
MOVJ C00329 VJ=10.00 ACC=20
MACRO1 MJ#(0) ARGF101
ARCON
MOVL C00330 V=13.5 ACC=20
ARCOF
TIMER T=7.00
*LABEL159
MOVJ C00331 VJ=10.00 ACC=20
MACRO1 MJ#(0) ARGF101
ARCON
MOVL C00332 V=13.5 ACC=20
ARCOF
DOUT OT#(9) ON
TIMER T=50.00
DOUT OT#(9) OFF
TIMER T=13.00
MOVJ C00333 VJ=10.00 ACC=20
*LABEL160
MOVJ C00334 VJ=10.00 ACC=20
MACRO1 MJ#(0) ARGF103
ARCON
MOVL C00335 V=13.5 ACC=20
ARCOF
TIMER T=7.00
*LABEL161
MOVJ C00336 VJ=10.00 ACC=20
MACRO1 MJ#(0) ARGF103
ARCON
MOVL C00337 V=13.5 ACC=20
ARCOF
TIMER T=7.00
*LABEL162
MOVJ C00338 VJ=10.00 ACC=20
MACRO1 MJ#(0) ARGF101
ARCON
MOVL C00339 V=13.5 ACC=20
ARCOF
TIMER T=7.00
*LABEL163
MOVJ C00340 VJ=10.00 ACC=20
MACRO1 MJ#(0) ARGF101
ARCON
MOVL C00341 V=13.5 ACC=20
ARCOF
TIMER T=7.00
*LABEL164
MOVJ C00342 VJ=10.00 ACC=20
MACRO1 MJ#(0) ARGF101
ARCON
MOVL C00343 V=13.5 ACC=20
ARCOF
TIMER T=7.00
*LABEL165
MOVJ C00344 VJ=10.00 ACC=20
MACRO1 MJ#(0) ARGF101
ARCON
MOVL C00345 V=13.5 ACC=20
ARCOF
TIMER T=7.00
*LABEL166
MOVJ C00346 VJ=10.00 ACC=20
MACRO1 MJ#(0) ARGF101
ARCON
MOVL C00347 V=13.5 ACC=20
ARCOF
TIMER T=7.00
*LABEL167
MOVJ C00348 VJ=10.00 ACC=20
MACRO1 MJ#(0) ARGF101
ARCON
MOVL C00349 V=13.5 ACC=20
ARCOF
TIMER T=7.00
*LABEL168
MOVJ C00350 VJ=10.00 ACC=20
MACRO1 MJ#(0) ARGF101
ARCON
MOVL C00351 V=13.5 ACC=20
ARCOF
TIMER T=7.00
*LABEL169
MOVJ C00352 VJ=10.00 ACC=20
MACRO1 MJ#(0) ARGF101
ARCON
MOVL C00353 V=13.5 ACC=20
ARCOF
TIMER T=7.00
*LABEL170
MOVJ C00354 VJ=10.00 ACC=20
MACRO1 MJ#(0) ARGF101
ARCON
MOVL C00355 V=13.5 ACC=20
ARCOF
TIMER T=7.00
*LABEL171
MOVJ C00356 VJ=10.00 ACC=20
MACRO1 MJ#(0) ARGF101
ARCON
MOVL C00357 V=13.5 ACC=20
ARCOF
DOUT OT#(9) ON
TIMER T=50.00
DOUT OT#(9) OFF
TIMER T=13.00
MOVJ C00358 VJ=10.00 ACC=20
*LABEL172
MOVJ C00359 VJ=10.00 ACC=20
MACRO1 MJ#(0) ARGF103
ARCON
MOVL C00360 V=13.5 ACC=20
ARCOF
TIMER T=7.00
*LABEL173
MOVJ C00361 VJ=10.00 ACC=20
MACRO1 MJ#(0) ARGF103
ARCON
MOVL C00362 V=13.5 ACC=20
ARCOF
TIMER T=7.00
*LABEL174
MOVJ C00363 VJ=10.00 ACC=20
MACRO1 MJ#(0) ARGF101
ARCON
MOVL C00364 V=13.5 ACC=20
ARCOF
TIMER T=7.00
*LABEL175
MOVJ C00365 VJ=10.00 ACC=20
MACRO1 MJ#(0) ARGF101
ARCON
MOVL C00366 V=13.5 ACC=20
ARCOF
TIMER T=7.00
*LABEL176
MOVJ C00367 VJ=10.00 ACC=20
MACRO1 MJ#(0) ARGF101
ARCON
MOVL C00368 V=13.5 ACC=20
ARCOF
TIMER T=7.00
*LABEL177
MOVJ C00369 VJ=10.00 ACC=20
MACRO1 MJ#(0) ARGF101
ARCON
MOVL C00370 V=13.5 ACC=20
ARCOF
TIMER T=7.00
*LABEL178
MOVJ C00371 VJ=10.00 ACC=20
MACRO1 MJ#(0) ARGF101
ARCON
MOVL C00372 V=13.5 ACC=20
ARCOF
TIMER T=7.00
*LABEL179
MOVJ C00373 VJ=10.00 ACC=20
MACRO1 MJ#(0) ARGF101
ARCON
MOVL C00374 V=13.5 ACC=20
ARCOF
TIMER T=7.00
*LABEL180
MOVJ C00375 VJ=10.00 ACC=20
MACRO1 MJ#(0) ARGF101
ARCON
MOVL C00376 V=13.5 ACC=20
ARCOF
TIMER T=7.00
*LABEL181
MOVJ C00377 VJ=10.00 ACC=20
MACRO1 MJ#(0) ARGF101
ARCON
MOVL C00378 V=13.5 ACC=20
ARCOF
TIMER T=7.00
*LABEL182
MOVJ C00379 VJ=10.00 ACC=20
MACRO1 MJ#(0) ARGF101
ARCON
MOVL C00380 V=13.5 ACC=20
ARCOF
TIMER T=7.00
*LABEL183
MOVJ C00381 VJ=10.00 ACC=20
MACRO1 MJ#(0) ARGF101
ARCON
MOVL C00382 V=13.5 ACC=20
ARCOF
TIMER T=7.00
*LABEL184
MOVJ C00383 VJ=10.00 ACC=20
MACRO1 MJ#(0) ARGF103
ARCON
MOVL C00384 V=13.5 ACC=20
ARCOF
TIMER T=7.00
*LABEL185
MOVJ C00385 VJ=10.00 ACC=20
MACRO1 MJ#(0) ARGF103
ARCON
MOVL C00386 V=13.5 ACC=20
ARCOF
DOUT OT#(9) ON
TIMER T=50.00
DOUT OT#(9) OFF
TIMER T=13.00
MOVJ C00387 VJ=10.00 ACC=20
*LABEL186
MOVJ C00388 VJ=10.00 ACC=20
MACRO1 MJ#(0) ARGF103
ARCON
MOVL C00389 V=13.5 ACC=20
ARCOF
TIMER T=7.00
*LABEL187
MOVJ C00390 VJ=10.00 ACC=20
MACRO1 MJ#(0) ARGF103
ARCON
MOVL C00391 V=13.5 ACC=20
ARCOF
TIMER T=7.00
*LABEL188
MOVJ C00392 VJ=10.00 ACC=20
MACRO1 MJ#(0) ARGF101
ARCON
MOVL C00393 V=13.5 ACC=20
ARCOF
TIMER T=7.00
*LABEL189
MOVJ C00394 VJ=10.00 ACC=20
MACRO1 MJ#(0) ARGF101
ARCON
MOVL C00395 V=13.5 ACC=20
ARCOF
TIMER T=7.00
*LABEL190
MOVJ C00396 VJ=10.00 ACC=20
MACRO1 MJ#(0) ARGF101
ARCON
MOVL C00397 V=13.5 ACC=20
ARCOF
TIMER T=7.00
*LABEL191
MOVJ C00398 VJ=10.00 ACC=20
MACRO1 MJ#(0) ARGF101
ARCON
MOVL C00399 V=13.5 ACC=20
ARCOF
TIMER T=7.00
*LABEL192
MOVJ C00400 VJ=10.00 ACC=20
MACRO1 MJ#(0) ARGF101
ARCON
MOVL C00401 V=13.5 ACC=20
ARCOF
TIMER T=7.00
*LABEL193
MOVJ C00402 VJ=10.00 ACC=20
MACRO1 MJ#(0) ARGF101
ARCON
MOVL C00403 V=13.5 ACC=20
ARCOF
TIMER T=7.00
*LABEL194
MOVJ C00404 VJ=10.00 ACC=20
MACRO1 MJ#(0) ARGF101
ARCON
MOVL C00405 V=13.5 ACC=20
ARCOF
TIMER T=7.00
*LABEL195
MOVJ C00406 VJ=10.00 ACC=20
MACRO1 MJ#(0) ARGF101
ARCON
MOVL C00407 V=13.5 ACC=20
ARCOF
TIMER T=7.00
*LABEL196
MOVJ C00408 VJ=10.00 ACC=20
MACRO1 MJ#(0) ARGF101
ARCON
MOVL C00409 V=13.5 ACC=20
ARCOF
TIMER T=7.00
*LABEL197
MOVJ C00410 VJ=10.00 ACC=20
MACRO1 MJ#(0) ARGF101
ARCON
MOVL C00411 V=13.5 ACC=20
ARCOF
DOUT OT#(9) ON
TIMER T=50.00
DOUT OT#(9) OFF
TIMER T=13.00
MOVJ C00412 VJ=10.00 ACC=20
*LABEL198
MOVJ C00413 VJ=10.00 ACC=20
MACRO1 MJ#(0) ARGF103
ARCON
MOVL C00414 V=13.5 ACC=20
ARCOF
TIMER T=7.00
*LABEL199
MOVJ C00415 VJ=10.00 ACC=20
MACRO1 MJ#(0) ARGF103
ARCON
MOVL C00416 V=13.5 ACC=20
ARCOF
TIMER T=7.00
*LABEL200
MOVJ C00417 VJ=10.00 ACC=20
MACRO1 MJ#(0) ARGF101
ARCON
MOVL C00418 V=13.5 ACC=20
ARCOF
TIMER T=7.00
*LABEL201
MOVJ C00419 VJ=10.00 ACC=20
MACRO1 MJ#(0) ARGF101
ARCON
MOVL C00420 V=13.5 ACC=20
ARCOF
TIMER T=7.00
*LABEL202
MOVJ C00421 VJ=10.00 ACC=20
MACRO1 MJ#(0) ARGF101
ARCON
MOVL C00422 V=13.5 ACC=20
ARCOF
TIMER T=7.00
*LABEL203
MOVJ C00423 VJ=10.00 ACC=20
MACRO1 MJ#(0) ARGF101
ARCON
MOVL C00424 V=13.5 ACC=20
ARCOF
TIMER T=7.00
*LABEL204
MOVJ C00425 VJ=10.00 ACC=20
MACRO1 MJ#(0) ARGF101
ARCON
MOVL C00426 V=13.5 ACC=20
ARCOF
TIMER T=7.00
*LABEL205
MOVJ C00427 VJ=10.00 ACC=20
MACRO1 MJ#(0) ARGF101
ARCON
MOVL C00428 V=13.5 ACC=20
ARCOF
TIMER T=7.00
*LABEL206
MOVJ C00429 VJ=10.00 ACC=20
MACRO1 MJ#(0) ARGF101
ARCON
MOVL C00430 V=13.5 ACC=20
ARCOF
TIMER T=7.00
*LABEL207
MOVJ C00431 VJ=10.00 ACC=20
MACRO1 MJ#(0) ARGF101
ARCON
MOVL C00432 V=13.5 ACC=20
ARCOF
TIMER T=7.00
*LABEL208
MOVJ C00433 VJ=10.00 ACC=20
MACRO1 MJ#(0) ARGF101
ARCON
MOVL C00434 V=13.5 ACC=20
ARCOF
TIMER T=7.00
*LABEL209
MOVJ C00435 VJ=10.00 ACC=20
MACRO1 MJ#(0) ARGF101
ARCON
MOVL C00436 V=13.5 ACC=20
ARCOF
DOUT OT#(9) ON
TIMER T=50.00
DOUT OT#(9) OFF
TIMER T=13.00
MOVJ C00437 VJ=10.00 ACC=20
*LABEL210
MOVJ C00438 VJ=10.00 ACC=20
MACRO1 MJ#(0) ARGF103
ARCON
MOVL C00439 V=13.5 ACC=20
ARCOF
TIMER T=7.00
*LABEL211
MOVJ C00440 VJ=10.00 ACC=20
MACRO1 MJ#(0) ARGF103
ARCON
MOVL C00441 V=13.5 ACC=20
ARCOF
TIMER T=7.00
*LABEL212
MOVJ C00442 VJ=10.00 ACC=20
MACRO1 MJ#(0) ARGF101
ARCON
MOVL C00443 V=13.5 ACC=20
ARCOF
TIMER T=7.00
*LABEL213
MOVJ C00444 VJ=10.00 ACC=20
MACRO1 MJ#(0) ARGF101
ARCON
MOVL C00445 V=13.5 ACC=20
ARCOF
TIMER T=7.00
*LABEL214
MOVJ C00446 VJ=10.00 ACC=20
MACRO1 MJ#(0) ARGF101
ARCON
MOVL C00447 V=13.5 ACC=20
ARCOF
TIMER T=7.00
*LABEL215
MOVJ C00448 VJ=10.00 ACC=20
MACRO1 MJ#(0) ARGF101
ARCON
MOVL C00449 V=13.5 ACC=20
ARCOF
TIMER T=7.00
*LABEL216
MOVJ C00450 VJ=10.00 ACC=20
MACRO1 MJ#(0) ARGF101
ARCON
MOVL C00451 V=13.5 ACC=20
ARCOF
TIMER T=7.00
*LABEL217
MOVJ C00452 VJ=10.00 ACC=20
MACRO1 MJ#(0) ARGF101
ARCON
MOVL C00453 V=13.5 ACC=20
ARCOF
TIMER T=7.00
*LABEL218
MOVJ C00454 VJ=10.00 ACC=20
MACRO1 MJ#(0) ARGF101
ARCON
MOVL C00455 V=13.5 ACC=20
ARCOF
TIMER T=7.00
*LABEL219
MOVJ C00456 VJ=10.00 ACC=20
MACRO1 MJ#(0) ARGF101
ARCON
MOVL C00457 V=13.5 ACC=20
ARCOF
TIMER T=7.00
*LABEL220
MOVJ C00458 VJ=10.00 ACC=20
MACRO1 MJ#(0) ARGF101
ARCON
MOVL C00459 V=13.5 ACC=20
ARCOF
TIMER T=7.00
*LABEL221
MOVJ C00460 VJ=10.00 ACC=20
MACRO1 MJ#(0) ARGF101
ARCON
MOVL C00461 V=13.5 ACC=20
ARCOF
DOUT OT#(9) ON
TIMER T=50.00
DOUT OT#(9) OFF
TIMER T=13.00
MOVJ C00462 VJ=10.00 ACC=20
*LABEL222
MOVJ C00463 VJ=10.00 ACC=20
MACRO1 MJ#(0) ARGF103
ARCON
MOVL C00464 V=13.5 ACC=20
ARCOF
TIMER T=7.00
*LABEL223
MOVJ C00465 VJ=10.00 ACC=20
MACRO1 MJ#(0) ARGF103
ARCON
MOVL C00466 V=13.5 ACC=20
ARCOF
TIMER T=7.00
*LABEL224
MOVJ C00467 VJ=10.00 ACC=20
MACRO1 MJ#(0) ARGF101
ARCON
MOVL C00468 V=13.5 ACC=20
ARCOF
TIMER T=7.00
*LABEL225
MOVJ C00469 VJ=10.00 ACC=20
MACRO1 MJ#(0) ARGF101
ARCON
MOVL C00470 V=13.5 ACC=20
ARCOF
TIMER T=7.00
*LABEL226
MOVJ C00471 VJ=10.00 ACC=20
MACRO1 MJ#(0) ARGF101
ARCON
MOVL C00472 V=13.5 ACC=20
ARCOF
TIMER T=7.00
*LABEL227
MOVJ C00473 VJ=10.00 ACC=20
MACRO1 MJ#(0) ARGF101
ARCON
MOVL C00474 V=13.5 ACC=20
ARCOF
TIMER T=7.00
*LABEL228
MOVJ C00475 VJ=10.00 ACC=20
MACRO1 MJ#(0) ARGF101
ARCON
MOVL C00476 V=13.5 ACC=20
ARCOF
TIMER T=7.00
*LABEL229
MOVJ C00477 VJ=10.00 ACC=20
MACRO1 MJ#(0) ARGF101
ARCON
MOVL C00478 V=13.5 ACC=20
ARCOF
TIMER T=7.00
*LABEL230
MOVJ C00479 VJ=10.00 ACC=20
MACRO1 MJ#(0) ARGF101
ARCON
MOVL C00480 V=13.5 ACC=20
ARCOF
TIMER T=7.00
*LABEL231
MOVJ C00481 VJ=10.00 ACC=20
MACRO1 MJ#(0) ARGF101
ARCON
MOVL C00482 V=13.5 ACC=20
ARCOF
TIMER T=7.00
*LABEL232
MOVJ C00483 VJ=10.00 ACC=20
MACRO1 MJ#(0) ARGF101
ARCON
MOVL C00484 V=13.5 ACC=20
ARCOF
TIMER T=7.00
*LABEL233
MOVJ C00485 VJ=10.00 ACC=20
MACRO1 MJ#(0) ARGF101
ARCON
MOVL C00486 V=13.5 ACC=20
ARCOF
DOUT OT#(9) ON
TIMER T=50.00
DOUT OT#(9) OFF
TIMER T=13.00
MOVJ C00487 VJ=10.00 ACC=20
*LABEL234
MOVJ C00488 VJ=10.00 ACC=20
MACRO1 MJ#(0) ARGF103
ARCON
MOVL C00489 V=13.5 ACC=20
ARCOF
TIMER T=7.00
*LABEL235
MOVJ C00490 VJ=10.00 ACC=20
MACRO1 MJ#(0) ARGF103
ARCON
MOVL C00491 V=13.5 ACC=20
ARCOF
TIMER T=7.00
*LABEL236
MOVJ C00492 VJ=10.00 ACC=20
MACRO1 MJ#(0) ARGF101
ARCON
MOVL C00493 V=13.5 ACC=20
ARCOF
TIMER T=7.00
*LABEL237
MOVJ C00494 VJ=10.00 ACC=20
MACRO1 MJ#(0) ARGF101
ARCON
MOVL C00495 V=13.5 ACC=20
ARCOF
TIMER T=7.00
*LABEL238
MOVJ C00496 VJ=10.00 ACC=20
MACRO1 MJ#(0) ARGF101
ARCON
MOVL C00497 V=13.5 ACC=20
ARCOF
TIMER T=7.00
*LABEL239
MOVJ C00498 VJ=10.00 ACC=20
MACRO1 MJ#(0) ARGF101
ARCON
MOVL C00499 V=13.5 ACC=20
ARCOF
TIMER T=7.00
*LABEL240
MOVJ C00500 VJ=10.00 ACC=20
MACRO1 MJ#(0) ARGF101
ARCON
MOVL C00501 V=13.5 ACC=20
ARCOF
TIMER T=7.00
*LABEL241
MOVJ C00502 VJ=10.00 ACC=20
MACRO1 MJ#(0) ARGF101
ARCON
MOVL C00503 V=13.5 ACC=20
ARCOF
TIMER T=7.00
*LABEL242
MOVJ C00504 VJ=10.00 ACC=20
MACRO1 MJ#(0) ARGF101
ARCON
MOVL C00505 V=13.5 ACC=20
ARCOF
TIMER T=7.00
*LABEL243
MOVJ C00506 VJ=10.00 ACC=20
MACRO1 MJ#(0) ARGF101
ARCON
MOVL C00507 V=13.5 ACC=20
ARCOF
TIMER T=7.00
*LABEL244
MOVJ C00508 VJ=10.00 ACC=20
MACRO1 MJ#(0) ARGF101
ARCON
MOVL C00509 V=13.5 ACC=20
ARCOF
TIMER T=7.00
*LABEL245
MOVJ C00510 VJ=10.00 ACC=20
MACRO1 MJ#(0) ARGF101
ARCON
MOVL C00511 V=13.5 ACC=20
ARCOF
TIMER T=7.00
*LABEL246
MOVJ C00512 VJ=10.00 ACC=20
MACRO1 MJ#(0) ARGF103
ARCON
MOVL C00513 V=13.5 ACC=20
ARCOF
TIMER T=7.00
*LABEL247
MOVJ C00514 VJ=10.00 ACC=20
MACRO1 MJ#(0) ARGF103
ARCON
MOVL C00515 V=13.5 ACC=20
ARCOF
DOUT OT#(9) ON
TIMER T=50.00
DOUT OT#(9) OFF
TIMER T=13.00
MOVJ C00516 VJ=10.00 ACC=20
*LABEL248
MOVJ C00517 VJ=10.00 ACC=20
MACRO1 MJ#(0) ARGF103
ARCON
MOVL C00518 V=13.5 ACC=20
ARCOF
TIMER T=7.00
*LABEL249
MOVJ C00519 VJ=10.00 ACC=20
MACRO1 MJ#(0) ARGF103
ARCON
MOVL C00520 V=13.5 ACC=20
ARCOF
TIMER T=7.00
*LABEL250
MOVJ C00521 VJ=10.00 ACC=20
MACRO1 MJ#(0) ARGF101
ARCON
MOVL C00522 V=13.5 ACC=20
ARCOF
TIMER T=7.00
*LABEL251
MOVJ C00523 VJ=10.00 ACC=20
MACRO1 MJ#(0) ARGF101
ARCON
MOVL C00524 V=13.5 ACC=20
ARCOF
TIMER T=7.00
*LABEL252
MOVJ C00525 VJ=10.00 ACC=20
MACRO1 MJ#(0) ARGF101
ARCON
MOVL C00526 V=13.5 ACC=20
ARCOF
TIMER T=7.00
*LABEL253
MOVJ C00527 VJ=10.00 ACC=20
MACRO1 MJ#(0) ARGF101
ARCON
MOVL C00528 V=13.5 ACC=20
ARCOF
TIMER T=7.00
*LABEL254
MOVJ C00529 VJ=10.00 ACC=20
MACRO1 MJ#(0) ARGF101
ARCON
MOVL C00530 V=13.5 ACC=20
ARCOF
TIMER T=7.00
*LABEL255
MOVJ C00531 VJ=10.00 ACC=20
MACRO1 MJ#(0) ARGF101
ARCON
MOVL C00532 V=13.5 ACC=20
ARCOF
TIMER T=7.00
*LABEL256
MOVJ C00533 VJ=10.00 ACC=20
MACRO1 MJ#(0) ARGF101
ARCON
MOVL C00534 V=13.5 ACC=20
ARCOF
TIMER T=7.00
*LABEL257
MOVJ C00535 VJ=10.00 ACC=20
MACRO1 MJ#(0) ARGF101
ARCON
MOVL C00536 V=13.5 ACC=20
ARCOF
TIMER T=7.00
*LABEL258
MOVJ C00537 VJ=10.00 ACC=20
MACRO1 MJ#(0) ARGF101
ARCON
MOVL C00538 V=13.5 ACC=20
ARCOF
TIMER T=7.00
*LABEL259
MOVJ C00539 VJ=10.00 ACC=20
MACRO1 MJ#(0) ARGF101
ARCON
MOVL C00540 V=13.5 ACC=20
ARCOF
DOUT OT#(9) ON
TIMER T=50.00
DOUT OT#(9) OFF
TIMER T=13.00
MOVJ C00541 VJ=10.00 ACC=20
*LABEL260
MOVJ C00542 VJ=10.00 ACC=20
MACRO1 MJ#(0) ARGF103
ARCON
MOVL C00543 V=13.5 ACC=20
ARCOF
TIMER T=7.00
*LABEL261
MOVJ C00544 VJ=10.00 ACC=20
MACRO1 MJ#(0) ARGF103
ARCON
MOVL C00545 V=13.5 ACC=20
ARCOF
TIMER T=7.00
*LABEL262
MOVJ C00546 VJ=10.00 ACC=20
MACRO1 MJ#(0) ARGF101
ARCON
MOVL C00547 V=13.5 ACC=20
ARCOF
TIMER T=7.00
*LABEL263
MOVJ C00548 VJ=10.00 ACC=20
MACRO1 MJ#(0) ARGF101
ARCON
MOVL C00549 V=13.5 ACC=20
ARCOF
TIMER T=7.00
*LABEL264
MOVJ C00550 VJ=10.00 ACC=20
MACRO1 MJ#(0) ARGF101
ARCON
MOVL C00551 V=13.5 ACC=20
ARCOF
TIMER T=7.00
*LABEL265
MOVJ C00552 VJ=10.00 ACC=20
MACRO1 MJ#(0) ARGF101
ARCON
MOVL C00553 V=13.5 ACC=20
ARCOF
TIMER T=7.00
*LABEL266
MOVJ C00554 VJ=10.00 ACC=20
MACRO1 MJ#(0) ARGF101
ARCON
MOVL C00555 V=13.5 ACC=20
ARCOF
TIMER T=7.00
*LABEL267
MOVJ C00556 VJ=10.00 ACC=20
MACRO1 MJ#(0) ARGF101
ARCON
MOVL C00557 V=13.5 ACC=20
ARCOF
TIMER T=7.00
*LABEL268
MOVJ C00558 VJ=10.00 ACC=20
MACRO1 MJ#(0) ARGF101
ARCON
MOVL C00559 V=13.5 ACC=20
ARCOF
TIMER T=7.00
*LABEL269
MOVJ C00560 VJ=10.00 ACC=20
MACRO1 MJ#(0) ARGF101
ARCON
MOVL C00561 V=13.5 ACC=20
ARCOF
TIMER T=7.00
*LABEL270
MOVJ C00562 VJ=10.00 ACC=20
MACRO1 MJ#(0) ARGF101
ARCON
MOVL C00563 V=13.5 ACC=20
ARCOF
TIMER T=7.00
*LABEL271
MOVJ C00564 VJ=10.00 ACC=20
MACRO1 MJ#(0) ARGF101
ARCON
MOVL C00565 V=13.5 ACC=20
ARCOF
DOUT OT#(9) ON
TIMER T=50.00
DOUT OT#(9) OFF
TIMER T=13.00
MOVJ C00566 VJ=10.00 ACC=20
*LABEL272
MOVJ C00567 VJ=10.00 ACC=20
MACRO1 MJ#(0) ARGF103
ARCON
MOVL C00568 V=13.5 ACC=20
ARCOF
TIMER T=7.00
*LABEL273
MOVJ C00569 VJ=10.00 ACC=20
MACRO1 MJ#(0) ARGF103
ARCON
MOVL C00570 V=13.5 ACC=20
ARCOF
TIMER T=7.00
*LABEL274
MOVJ C00571 VJ=10.00 ACC=20
MACRO1 MJ#(0) ARGF101
ARCON
MOVL C00572 V=13.5 ACC=20
ARCOF
TIMER T=7.00
*LABEL275
MOVJ C00573 VJ=10.00 ACC=20
MACRO1 MJ#(0) ARGF101
ARCON
MOVL C00574 V=13.5 ACC=20
ARCOF
TIMER T=7.00
*LABEL276
MOVJ C00575 VJ=10.00 ACC=20
MACRO1 MJ#(0) ARGF101
ARCON
MOVL C00576 V=13.5 ACC=20
ARCOF
TIMER T=7.00
*LABEL277
MOVJ C00577 VJ=10.00 ACC=20
MACRO1 MJ#(0) ARGF101
ARCON
MOVL C00578 V=13.5 ACC=20
ARCOF
TIMER T=7.00
*LABEL278
MOVJ C00579 VJ=10.00 ACC=20
MACRO1 MJ#(0) ARGF101
ARCON
MOVL C00580 V=13.5 ACC=20
ARCOF
TIMER T=7.00
*LABEL279
MOVJ C00581 VJ=10.00 ACC=20
MACRO1 MJ#(0) ARGF101
ARCON
MOVL C00582 V=13.5 ACC=20
ARCOF
TIMER T=7.00
*LABEL280
MOVJ C00583 VJ=10.00 ACC=20
MACRO1 MJ#(0) ARGF101
ARCON
MOVL C00584 V=13.5 ACC=20
ARCOF
TIMER T=7.00
*LABEL281
MOVJ C00585 VJ=10.00 ACC=20
MACRO1 MJ#(0) ARGF101
ARCON
MOVL C00586 V=13.5 ACC=20
ARCOF
TIMER T=7.00
*LABEL282
MOVJ C00587 VJ=10.00 ACC=20
MACRO1 MJ#(0) ARGF101
ARCON
MOVL C00588 V=13.5 ACC=20
ARCOF
TIMER T=7.00
*LABEL283
MOVJ C00589 VJ=10.00 ACC=20
MACRO1 MJ#(0) ARGF101
ARCON
MOVL C00590 V=13.5 ACC=20
ARCOF
DOUT OT#(9) ON
TIMER T=50.00
DOUT OT#(9) OFF
TIMER T=13.00
MOVJ C00591 VJ=10.00 ACC=20
*LABEL284
MOVJ C00592 VJ=10.00 ACC=20
MACRO1 MJ#(0) ARGF103
ARCON
MOVL C00593 V=13.5 ACC=20
ARCOF
TIMER T=7.00
*LABEL285
MOVJ C00594 VJ=10.00 ACC=20
MACRO1 MJ#(0) ARGF103
ARCON
MOVL C00595 V=13.5 ACC=20
ARCOF
TIMER T=7.00
*LABEL286
MOVJ C00596 VJ=10.00 ACC=20
MACRO1 MJ#(0) ARGF101
ARCON
MOVL C00597 V=13.5 ACC=20
ARCOF
TIMER T=7.00
*LABEL287
MOVJ C00598 VJ=10.00 ACC=20
MACRO1 MJ#(0) ARGF101
ARCON
MOVL C00599 V=13.5 ACC=20
ARCOF
TIMER T=7.00
*LABEL288
MOVJ C00600 VJ=10.00 ACC=20
MACRO1 MJ#(0) ARGF101
ARCON
MOVL C00601 V=13.5 ACC=20
ARCOF
TIMER T=7.00
*LABEL289
MOVJ C00602 VJ=10.00 ACC=20
MACRO1 MJ#(0) ARGF101
ARCON
MOVL C00603 V=13.5 ACC=20
ARCOF
TIMER T=7.00
*LABEL290
MOVJ C00604 VJ=10.00 ACC=20
MACRO1 MJ#(0) ARGF101
ARCON
MOVL C00605 V=13.5 ACC=20
ARCOF
TIMER T=7.00
*LABEL291
MOVJ C00606 VJ=10.00 ACC=20
MACRO1 MJ#(0) ARGF101
ARCON
MOVL C00607 V=13.5 ACC=20
ARCOF
TIMER T=7.00
*LABEL292
MOVJ C00608 VJ=10.00 ACC=20
MACRO1 MJ#(0) ARGF101
ARCON
MOVL C00609 V=13.5 ACC=20
ARCOF
TIMER T=7.00
*LABEL293
MOVJ C00610 VJ=10.00 ACC=20
MACRO1 MJ#(0) ARGF101
ARCON
MOVL C00611 V=13.5 ACC=20
ARCOF
TIMER T=7.00
*LABEL294
MOVJ C00612 VJ=10.00 ACC=20
MACRO1 MJ#(0) ARGF101
ARCON
MOVL C00613 V=13.5 ACC=20
ARCOF
TIMER T=7.00
*LABEL295
MOVJ C00614 VJ=10.00 ACC=20
MACRO1 MJ#(0) ARGF101
ARCON
MOVL C00615 V=13.5 ACC=20
ARCOF
DOUT OT#(9) ON
TIMER T=50.00
DOUT OT#(9) OFF
TIMER T=13.00
MOVJ C00616 VJ=10.00 ACC=20
*LABEL296
MOVJ C00617 VJ=10.00 ACC=20
MACRO1 MJ#(0) ARGF103
ARCON
MOVL C00618 V=13.5 ACC=20
ARCOF
TIMER T=7.00
*LABEL297
MOVJ C00619 VJ=10.00 ACC=20
MACRO1 MJ#(0) ARGF103
ARCON
MOVL C00620 V=13.5 ACC=20
ARCOF
TIMER T=7.00
*LABEL298
MOVJ C00621 VJ=10.00 ACC=20
MACRO1 MJ#(0) ARGF101
ARCON
MOVL C00622 V=13.5 ACC=20
ARCOF
TIMER T=7.00
*LABEL299
MOVJ C00623 VJ=10.00 ACC=20
MACRO1 MJ#(0) ARGF101
ARCON
MOVL C00624 V=13.5 ACC=20
ARCOF
TIMER T=7.00
*LABEL300
MOVJ C00625 VJ=10.00 ACC=20
MACRO1 MJ#(0) ARGF101
ARCON
MOVL C00626 V=13.5 ACC=20
ARCOF
TIMER T=7.00
*LABEL301
MOVJ C00627 VJ=10.00 ACC=20
MACRO1 MJ#(0) ARGF101
ARCON
MOVL C00628 V=13.5 ACC=20
ARCOF
TIMER T=7.00
*LABEL302
MOVJ C00629 VJ=10.00 ACC=20
MACRO1 MJ#(0) ARGF101
ARCON
MOVL C00630 V=13.5 ACC=20
ARCOF
TIMER T=7.00
*LABEL303
MOVJ C00631 VJ=10.00 ACC=20
MACRO1 MJ#(0) ARGF101
ARCON
MOVL C00632 V=13.5 ACC=20
ARCOF
TIMER T=7.00
*LABEL304
MOVJ C00633 VJ=10.00 ACC=20
MACRO1 MJ#(0) ARGF101
ARCON
MOVL C00634 V=13.5 ACC=20
ARCOF
TIMER T=7.00
*LABEL305
MOVJ C00635 VJ=10.00 ACC=20
MACRO1 MJ#(0) ARGF101
ARCON
MOVL C00636 V=13.5 ACC=20
ARCOF
TIMER T=7.00
*LABEL306
MOVJ C00637 VJ=10.00 ACC=20
MACRO1 MJ#(0) ARGF101
ARCON
MOVL C00638 V=13.5 ACC=20
ARCOF
TIMER T=7.00
*LABEL307
MOVJ C00639 VJ=10.00 ACC=20
MACRO1 MJ#(0) ARGF101
ARCON
MOVL C00640 V=13.5 ACC=20
ARCOF
TIMER T=7.00
*LABEL308
MOVJ C00641 VJ=10.00 ACC=20
MACRO1 MJ#(0) ARGF103
ARCON
MOVL C00642 V=13.5 ACC=20
ARCOF
TIMER T=7.00
*LABEL309
MOVJ C00643 VJ=10.00 ACC=20
MACRO1 MJ#(0) ARGF103
ARCON
MOVL C00644 V=13.5 ACC=20
ARCOF
DOUT OT#(9) ON
TIMER T=50.00
DOUT OT#(9) OFF
TIMER T=13.00
MOVJ C00645 VJ=10.00 ACC=20
*LABEL310
MOVJ C00646 VJ=10.00 ACC=20
MACRO1 MJ#(0) ARGF103
ARCON
MOVL C00647 V=13.5 ACC=20
ARCOF
TIMER T=7.00
*LABEL311
MOVJ C00648 VJ=10.00 ACC=20
MACRO1 MJ#(0) ARGF103
ARCON
MOVL C00649 V=13.5 ACC=20
ARCOF
TIMER T=7.00
*LABEL312
MOVJ C00650 VJ=10.00 ACC=20
MACRO1 MJ#(0) ARGF101
ARCON
MOVL C00651 V=13.5 ACC=20
ARCOF
TIMER T=7.00
*LABEL313
MOVJ C00652 VJ=10.00 ACC=20
MACRO1 MJ#(0) ARGF101
ARCON
MOVL C00653 V=13.5 ACC=20
ARCOF
TIMER T=7.00
*LABEL314
MOVJ C00654 VJ=10.00 ACC=20
MACRO1 MJ#(0) ARGF101
ARCON
MOVL C00655 V=13.5 ACC=20
ARCOF
TIMER T=7.00
*LABEL315
MOVJ C00656 VJ=10.00 ACC=20
MACRO1 MJ#(0) ARGF101
ARCON
MOVL C00657 V=13.5 ACC=20
ARCOF
TIMER T=7.00
*LABEL316
MOVJ C00658 VJ=10.00 ACC=20
MACRO1 MJ#(0) ARGF101
ARCON
MOVL C00659 V=13.5 ACC=20
ARCOF
TIMER T=7.00
*LABEL317
MOVJ C00660 VJ=10.00 ACC=20
MACRO1 MJ#(0) ARGF101
ARCON
MOVL C00661 V=13.5 ACC=20
ARCOF
TIMER T=7.00
*LABEL318
MOVJ C00662 VJ=10.00 ACC=20
MACRO1 MJ#(0) ARGF101
ARCON
MOVL C00663 V=13.5 ACC=20
ARCOF
TIMER T=7.00
*LABEL319
MOVJ C00664 VJ=10.00 ACC=20
MACRO1 MJ#(0) ARGF101
ARCON
MOVL C00665 V=13.5 ACC=20
ARCOF
TIMER T=7.00
*LABEL320
MOVJ C00666 VJ=10.00 ACC=20
MACRO1 MJ#(0) ARGF101
ARCON
MOVL C00667 V=13.5 ACC=20
ARCOF
TIMER T=7.00
*LABEL321
MOVJ C00668 VJ=10.00 ACC=20
MACRO1 MJ#(0) ARGF101
ARCON
MOVL C00669 V=13.5 ACC=20
ARCOF
DOUT OT#(9) ON
TIMER T=50.00
DOUT OT#(9) OFF
TIMER T=13.00
MOVJ C00670 VJ=10.00 ACC=20
*LABEL322
MOVJ C00671 VJ=10.00 ACC=20
MACRO1 MJ#(0) ARGF103
ARCON
MOVL C00672 V=13.5 ACC=20
ARCOF
TIMER T=7.00
*LABEL323
MOVJ C00673 VJ=10.00 ACC=20
MACRO1 MJ#(0) ARGF103
ARCON
MOVL C00674 V=13.5 ACC=20
ARCOF
TIMER T=7.00
*LABEL324
MOVJ C00675 VJ=10.00 ACC=20
MACRO1 MJ#(0) ARGF101
ARCON
MOVL C00676 V=13.5 ACC=20
ARCOF
TIMER T=7.00
*LABEL325
MOVJ C00677 VJ=10.00 ACC=20
MACRO1 MJ#(0) ARGF101
ARCON
MOVL C00678 V=13.5 ACC=20
ARCOF
TIMER T=7.00
*LABEL326
MOVJ C00679 VJ=10.00 ACC=20
MACRO1 MJ#(0) ARGF101
ARCON
MOVL C00680 V=13.5 ACC=20
ARCOF
TIMER T=7.00
*LABEL327
MOVJ C00681 VJ=10.00 ACC=20
MACRO1 MJ#(0) ARGF101
ARCON
MOVL C00682 V=13.5 ACC=20
ARCOF
TIMER T=7.00
*LABEL328
MOVJ C00683 VJ=10.00 ACC=20
MACRO1 MJ#(0) ARGF101
ARCON
MOVL C00684 V=13.5 ACC=20
ARCOF
TIMER T=7.00
*LABEL329
MOVJ C00685 VJ=10.00 ACC=20
MACRO1 MJ#(0) ARGF101
ARCON
MOVL C00686 V=13.5 ACC=20
ARCOF
TIMER T=7.00
*LABEL330
MOVJ C00687 VJ=10.00 ACC=20
MACRO1 MJ#(0) ARGF101
ARCON
MOVL C00688 V=13.5 ACC=20
ARCOF
TIMER T=7.00
*LABEL331
MOVJ C00689 VJ=10.00 ACC=20
MACRO1 MJ#(0) ARGF101
ARCON
MOVL C00690 V=13.5 ACC=20
ARCOF
TIMER T=7.00
*LABEL332
MOVJ C00691 VJ=10.00 ACC=20
MACRO1 MJ#(0) ARGF101
ARCON
MOVL C00692 V=13.5 ACC=20
ARCOF
TIMER T=7.00
*LABEL333
MOVJ C00693 VJ=10.00 ACC=20
MACRO1 MJ#(0) ARGF101
ARCON
MOVL C00694 V=13.5 ACC=20
ARCOF
DOUT OT#(9) ON
TIMER T=50.00
DOUT OT#(9) OFF
TIMER T=13.00
MOVJ C00695 VJ=10.00 ACC=20
*LABEL334
MOVJ C00696 VJ=10.00 ACC=20
MACRO1 MJ#(0) ARGF103
ARCON
MOVL C00697 V=13.5 ACC=20
ARCOF
TIMER T=7.00
*LABEL335
MOVJ C00698 VJ=10.00 ACC=20
MACRO1 MJ#(0) ARGF103
ARCON
MOVL C00699 V=13.5 ACC=20
ARCOF
TIMER T=7.00
*LABEL336
MOVJ C00700 VJ=10.00 ACC=20
MACRO1 MJ#(0) ARGF101
ARCON
MOVL C00701 V=13.5 ACC=20
ARCOF
TIMER T=7.00
*LABEL337
MOVJ C00702 VJ=10.00 ACC=20
MACRO1 MJ#(0) ARGF101
ARCON
MOVL C00703 V=13.5 ACC=20
ARCOF
TIMER T=7.00
*LABEL338
MOVJ C00704 VJ=10.00 ACC=20
MACRO1 MJ#(0) ARGF101
ARCON
MOVL C00705 V=13.5 ACC=20
ARCOF
TIMER T=7.00
*LABEL339
MOVJ C00706 VJ=10.00 ACC=20
MACRO1 MJ#(0) ARGF101
ARCON
MOVL C00707 V=13.5 ACC=20
ARCOF
TIMER T=7.00
*LABEL340
MOVJ C00708 VJ=10.00 ACC=20
MACRO1 MJ#(0) ARGF101
ARCON
MOVL C00709 V=13.5 ACC=20
ARCOF
TIMER T=7.00
*LABEL341
MOVJ C00710 VJ=10.00 ACC=20
MACRO1 MJ#(0) ARGF101
ARCON
MOVL C00711 V=13.5 ACC=20
ARCOF
TIMER T=7.00
*LABEL342
MOVJ C00712 VJ=10.00 ACC=20
MACRO1 MJ#(0) ARGF101
ARCON
MOVL C00713 V=13.5 ACC=20
ARCOF
TIMER T=7.00
*LABEL343
MOVJ C00714 VJ=10.00 ACC=20
MACRO1 MJ#(0) ARGF101
ARCON
MOVL C00715 V=13.5 ACC=20
ARCOF
TIMER T=7.00
*LABEL344
MOVJ C00716 VJ=10.00 ACC=20
MACRO1 MJ#(0) ARGF101
ARCON
MOVL C00717 V=13.5 ACC=20
ARCOF
TIMER T=7.00
*LABEL345
MOVJ C00718 VJ=10.00 ACC=20
MACRO1 MJ#(0) ARGF101
ARCON
MOVL C00719 V=13.5 ACC=20
ARCOF
DOUT OT#(9) ON
TIMER T=50.00
DOUT OT#(9) OFF
TIMER T=13.00
MOVJ C00720 VJ=10.00 ACC=20
*LABEL346
MOVJ C00721 VJ=10.00 ACC=20
MACRO1 MJ#(0) ARGF103
ARCON
MOVL C00722 V=13.5 ACC=20
ARCOF
TIMER T=7.00
*LABEL347
MOVJ C00723 VJ=10.00 ACC=20
MACRO1 MJ#(0) ARGF103
ARCON
MOVL C00724 V=13.5 ACC=20
ARCOF
TIMER T=7.00
*LABEL348
MOVJ C00725 VJ=10.00 ACC=20
MACRO1 MJ#(0) ARGF101
ARCON
MOVL C00726 V=13.5 ACC=20
ARCOF
TIMER T=7.00
*LABEL349
MOVJ C00727 VJ=10.00 ACC=20
MACRO1 MJ#(0) ARGF101
ARCON
MOVL C00728 V=13.5 ACC=20
ARCOF
TIMER T=7.00
*LABEL350
MOVJ C00729 VJ=10.00 ACC=20
MACRO1 MJ#(0) ARGF101
ARCON
MOVL C00730 V=13.5 ACC=20
ARCOF
TIMER T=7.00
*LABEL351
MOVJ C00731 VJ=10.00 ACC=20
MACRO1 MJ#(0) ARGF101
ARCON
MOVL C00732 V=13.5 ACC=20
ARCOF
TIMER T=7.00
*LABEL352
MOVJ C00733 VJ=10.00 ACC=20
MACRO1 MJ#(0) ARGF101
ARCON
MOVL C00734 V=13.5 ACC=20
ARCOF
TIMER T=7.00
*LABEL353
MOVJ C00735 VJ=10.00 ACC=20
MACRO1 MJ#(0) ARGF101
ARCON
MOVL C00736 V=13.5 ACC=20
ARCOF
TIMER T=7.00
*LABEL354
MOVJ C00737 VJ=10.00 ACC=20
MACRO1 MJ#(0) ARGF101
ARCON
MOVL C00738 V=13.5 ACC=20
ARCOF
TIMER T=7.00
*LABEL355
MOVJ C00739 VJ=10.00 ACC=20
MACRO1 MJ#(0) ARGF101
ARCON
MOVL C00740 V=13.5 ACC=20
ARCOF
TIMER T=7.00
*LABEL356
MOVJ C00741 VJ=10.00 ACC=20
MACRO1 MJ#(0) ARGF101
ARCON
MOVL C00742 V=13.5 ACC=20
ARCOF
TIMER T=7.00
*LABEL357
MOVJ C00743 VJ=10.00 ACC=20
MACRO1 MJ#(0) ARGF101
ARCON
MOVL C00744 V=13.5 ACC=20
ARCOF
DOUT OT#(9) ON
TIMER T=50.00
DOUT OT#(9) OFF
TIMER T=13.00
MOVJ C00745 VJ=10.00 ACC=20
*LABEL358
MOVJ C00746 VJ=10.00 ACC=20
MACRO1 MJ#(0) ARGF103
ARCON
MOVL C00747 V=13.5 ACC=20
ARCOF
TIMER T=7.00
*LABEL359
MOVJ C00748 VJ=10.00 ACC=20
MACRO1 MJ#(0) ARGF103
ARCON
MOVL C00749 V=13.5 ACC=20
ARCOF
TIMER T=7.00
*LABEL360
MOVJ C00750 VJ=10.00 ACC=20
MACRO1 MJ#(0) ARGF101
ARCON
MOVL C00751 V=13.5 ACC=20
ARCOF
TIMER T=7.00
*LABEL361
MOVJ C00752 VJ=10.00 ACC=20
MACRO1 MJ#(0) ARGF101
ARCON
MOVL C00753 V=13.5 ACC=20
ARCOF
TIMER T=7.00
*LABEL362
MOVJ C00754 VJ=10.00 ACC=20
MACRO1 MJ#(0) ARGF101
ARCON
MOVL C00755 V=13.5 ACC=20
ARCOF
TIMER T=7.00
*LABEL363
MOVJ C00756 VJ=10.00 ACC=20
MACRO1 MJ#(0) ARGF101
ARCON
MOVL C00757 V=13.5 ACC=20
ARCOF
TIMER T=7.00
*LABEL364
MOVJ C00758 VJ=10.00 ACC=20
MACRO1 MJ#(0) ARGF101
ARCON
MOVL C00759 V=13.5 ACC=20
ARCOF
TIMER T=7.00
*LABEL365
MOVJ C00760 VJ=10.00 ACC=20
MACRO1 MJ#(0) ARGF101
ARCON
MOVL C00761 V=13.5 ACC=20
ARCOF
TIMER T=7.00
*LABEL366
MOVJ C00762 VJ=10.00 ACC=20
MACRO1 MJ#(0) ARGF101
ARCON
MOVL C00763 V=13.5 ACC=20
ARCOF
TIMER T=7.00
*LABEL367
MOVJ C00764 VJ=10.00 ACC=20
MACRO1 MJ#(0) ARGF101
ARCON
MOVL C00765 V=13.5 ACC=20
ARCOF
TIMER T=7.00
*LABEL368
MOVJ C00766 VJ=10.00 ACC=20
MACRO1 MJ#(0) ARGF101
ARCON
MOVL C00767 V=13.5 ACC=20
ARCOF
TIMER T=7.00
*LABEL369
MOVJ C00768 VJ=10.00 ACC=20
MACRO1 MJ#(0) ARGF101
ARCON
MOVL C00769 V=13.5 ACC=20
ARCOF
TIMER T=7.00
*LABEL370
MOVJ C00770 VJ=10.00 ACC=20
MACRO1 MJ#(0) ARGF103
ARCON
MOVL C00771 V=13.5 ACC=20
ARCOF
TIMER T=7.00
*LABEL371
MOVJ C00772 VJ=10.00 ACC=20
MACRO1 MJ#(0) ARGF103
ARCON
MOVL C00773 V=13.5 ACC=20
ARCOF
DOUT OT#(9) ON
TIMER T=50.00
DOUT OT#(9) OFF
TIMER T=13.00
MOVJ C00774 VJ=10.00 ACC=20
END
